    IF _runOneStep THEN
        _runOneStep := FALSE;
        RETURN;
    END_IF
END_IF

IF SUPER^.Step(765, TRUE, 'Step number 765') THEN
    SUPER^.StepCompleteWhen((_runOneStep OR _runAllSteps) AND _finishStep);

    IF _runOneStep THEN
        _runOneStep := FALSE;
        RETURN;
    END_IF
END_IF

IF SUPER^.Step(766, TRUE, 'Step number 766') THEN
    SUPER^.StepCompleteWhen((_runOneStep OR _runAllSteps) AND _finishStep);

    IF _runOneStep THEN
        _runOneStep := FALSE;
        RETURN;
    END_IF
END_IF

IF SUPER^.Step(767, TRUE, 'Step number 767') THEN
    SUPER^.StepCompleteWhen((_runOneStep OR _runAllSteps) AND _finishStep);

    IF _runOneStep THEN
        _runOneStep := FALSE;
        RETURN;
    END_IF
END_IF

IF SUPER^.Step(768, TRUE, 'Step number 768') THEN
    SUPER^.StepCompleteWhen((_runOneStep OR _runAllSteps) AND _finishStep);

    IF _runOneStep THEN
        _runOneStep := FALSE;
        RETURN;
    END_IF
END_IF

IF SUPER^.Step(769, TRUE, 'Step number 769') THEN
    SUPER^.StepCompleteWhen((_runOneStep OR _runAllSteps) AND _finishStep);

    IF _runOneStep THEN
        _runOneStep := FALSE;
        RETURN;
    END_IF
END_IF

IF SUPER^.Step(770, TRUE, 'Step number 770') THEN
    SUPER^.StepCompleteWhen((_runOneStep OR _runAllSteps) AND _finishStep);

    IF _runOneStep THEN
        _runOneStep := FALSE;
        RETURN;
    END_IF
END_IF

IF SUPER^.Step(771, TRUE, 'Step number 771') THEN
    SUPER^.StepCompleteWhen((_runOneStep OR _runAllSteps) AND _finishStep);

    IF _runOneStep THEN
        _runOneStep := FALSE;
        RETURN;
    END_IF
END_IF

IF SUPER^.Step(772, TRUE, 'Step number 772') THEN
    SUPER^.StepCompleteWhen((_runOneStep OR _runAllSteps) AND _finishStep);

    IF _runOneStep THEN
        _runOneStep := FALSE;
        RETURN;
    END_IF
END_IF

IF SUPER^.Step(773, TRUE, 'Step number 773') THEN
    SUPER^.StepCompleteWhen((_runOneStep OR _runAllSteps) AND _finishStep);

    IF _runOneStep THEN
        _runOneStep := FALSE;
        RETURN;
    END_IF
END_IF

IF SUPER^.Step(774, TRUE, 'Step number 774') THEN
    SUPER^.StepCompleteWhen((_runOneStep OR _runAllSteps) AND _finishStep);

    IF _runOneStep THEN
        _runOneStep := FALSE;
        RETURN;
    END_IF
END_IF

IF SUPER^.Step(775, TRUE, 'Step number 775') THEN
    SUPER^.StepCompleteWhen((_runOneStep OR _runAllSteps) AND _finishStep);

    IF _runOneStep THEN
        _runOneStep := FALSE;
        RETURN;
    END_IF
END_IF

IF SUPER^.Step(776, TRUE, 'Step number 776') THEN
    SUPER^.StepCompleteWhen((_runOneStep OR _runAllSteps) AND _finishStep);

    IF _runOneStep THEN
        _runOneStep := FALSE;
        RETURN;
    END_IF
END_IF

IF SUPER^.Step(777, TRUE, 'Step number 777') THEN
    SUPER^.StepCompleteWhen((_runOneStep OR _runAllSteps) AND _finishStep);

    IF _runOneStep THEN
        _runOneStep := FALSE;
        RETURN;
    END_IF
END_IF

IF SUPER^.Step(778, TRUE, 'Step number 778') THEN
    SUPER^.StepCompleteWhen((_runOneStep OR _runAllSteps) AND _finishStep);

    IF _runOneStep THEN
        _runOneStep := FALSE;
        RETURN;
    END_IF
END_IF

IF SUPER^.Step(779, TRUE, 'Step number 779') THEN
    SUPER^.StepCompleteWhen((_runOneStep OR _runAllSteps) AND _finishStep);

    IF _runOneStep THEN
        _runOneStep := FALSE;
        RETURN;
    END_IF
END_IF

IF SUPER^.Step(780, TRUE, 'Step number 780') THEN
    SUPER^.StepCompleteWhen((_runOneStep OR _runAllSteps) AND _finishStep);

    IF _runOneStep THEN
        _runOneStep := FALSE;
        RETURN;
    END_IF
END_IF

IF SUPER^.Step(781, TRUE, 'Step number 781') THEN
    SUPER^.StepCompleteWhen((_runOneStep OR _runAllSteps) AND _finishStep);

    IF _runOneStep THEN
        _runOneStep := FALSE;
        RETURN;
    END_IF
END_IF

IF SUPER^.Step(782, TRUE, 'Step number 782') THEN
    SUPER^.StepCompleteWhen((_runOneStep OR _runAllSteps) AND _finishStep);

    IF _runOneStep THEN
        _runOneStep := FALSE;
        RETURN;
    END_IF
END_IF

IF SUPER^.Step(783, TRUE, 'Step number 783') THEN
    SUPER^.StepCompleteWhen((_runOneStep OR _runAllSteps) AND _finishStep);

    IF _runOneStep THEN
        _runOneStep := FALSE;
        RETURN;
    END_IF
END_IF

IF SUPER^.Step(784, TRUE, 'Step number 784') THEN
    SUPER^.StepCompleteWhen((_runOneStep OR _runAllSteps) AND _finishStep);

    IF _runOneStep THEN
        _runOneStep := FALSE;
        RETURN;
    END_IF
END_IF

IF SUPER^.Step(785, TRUE, 'Step number 785') THEN
    SUPER^.StepCompleteWhen((_runOneStep OR _runAllSteps) AND _finishStep);

    IF _runOneStep THEN
        _runOneStep := FALSE;
        RETURN;
    END_IF
END_IF

IF SUPER^.Step(786, TRUE, 'Step number 786') THEN
    SUPER^.StepCompleteWhen((_runOneStep OR _runAllSteps) AND _finishStep);

    IF _runOneStep THEN
        _runOneStep := FALSE;
        RETURN;
    END_IF
END_IF

IF SUPER^.Step(787, TRUE, 'Step number 787') THEN
    SUPER^.StepCompleteWhen((_runOneStep OR _runAllSteps) AND _finishStep);

    IF _runOneStep THEN
        _runOneStep := FALSE;
        RETURN;
    END_IF
END_IF

IF SUPER^.Step(788, TRUE, 'Step number 788') THEN
    SUPER^.StepCompleteWhen((_runOneStep OR _runAllSteps) AND _finishStep);

    IF _runOneStep THEN
        _runOneStep := FALSE;
        RETURN;
    END_IF
END_IF

IF SUPER^.Step(789, TRUE, 'Step number 789') THEN
    SUPER^.StepCompleteWhen((_runOneStep OR _runAllSteps) AND _finishStep);

    IF _runOneStep THEN
        _runOneStep := FALSE;
        RETURN;
    END_IF
END_IF

IF SUPER^.Step(790, TRUE, 'Step number 790') THEN
    SUPER^.StepCompleteWhen((_runOneStep OR _runAllSteps) AND _finishStep);

    IF _runOneStep THEN
        _runOneStep := FALSE;
        RETURN;
    END_IF
END_IF

IF SUPER^.Step(791, TRUE, 'Step number 791') THEN
    SUPER^.StepCompleteWhen((_runOneStep OR _runAllSteps) AND _finishStep);

    IF _runOneStep THEN
        _runOneStep := FALSE;
        RETURN;
    END_IF
END_IF

IF SUPER^.Step(792, TRUE, 'Step number 792') THEN
    SUPER^.StepCompleteWhen((_runOneStep OR _runAllSteps) AND _finishStep);

    IF _runOneStep THEN
        _runOneStep := FALSE;
        RETURN;
    END_IF
END_IF

IF SUPER^.Step(793, TRUE, 'Step number 793') THEN
    SUPER^.StepCompleteWhen((_runOneStep OR _runAllSteps) AND _finishStep);

    IF _runOneStep THEN
        _runOneStep := FALSE;
        RETURN;
    END_IF
END_IF

IF SUPER^.Step(794, TRUE, 'Step number 794') THEN
    SUPER^.StepCompleteWhen((_runOneStep OR _runAllSteps) AND _finishStep);

    IF _runOneStep THEN
        _runOneStep := FALSE;
        RETURN;
    END_IF
END_IF

IF SUPER^.Step(795, TRUE, 'Step number 795') THEN
    SUPER^.StepCompleteWhen((_runOneStep OR _runAllSteps) AND _finishStep);

    IF _runOneStep THEN
        _runOneStep := FALSE;
        RETURN;
    END_IF
END_IF

IF SUPER^.Step(796, TRUE, 'Step number 796') THEN
    SUPER^.StepCompleteWhen((_runOneStep OR _runAllSteps) AND _finishStep);

    IF _runOneStep THEN
        _runOneStep := FALSE;
        RETURN;
    END_IF
END_IF

IF SUPER^.Step(797, TRUE, 'Step number 797') THEN
    SUPER^.StepCompleteWhen((_runOneStep OR _runAllSteps) AND _finishStep);

    IF _runOneStep THEN
        _runOneStep := FALSE;
        RETURN;
    END_IF
END_IF

IF SUPER^.Step(798, TRUE, 'Step number 798') THEN
    SUPER^.StepCompleteWhen((_runOneStep OR _runAllSteps) AND _finishStep);

    IF _runOneStep THEN
        _runOneStep := FALSE;
        RETURN;
    END_IF
END_IF

IF SUPER^.Step(799, TRUE, 'Step number 799') THEN
    SUPER^.StepCompleteWhen((_runOneStep OR _runAllSteps) AND _finishStep);

    IF _runOneStep THEN
        _runOneStep := FALSE;
        RETURN;
    END_IF
END_IF

IF SUPER^.Step(800, TRUE, 'Step number 800') THEN
    SUPER^.StepCompleteWhen((_runOneStep OR _runAllSteps) AND _finishStep);

    IF _runOneStep THEN
        _runOneStep := FALSE;
        RETURN;
    END_IF
END_IF

IF SUPER^.Step(801, TRUE, 'Step number 801') THEN
    SUPER^.StepCompleteWhen((_runOneStep OR _runAllSteps) AND _finishStep);

    IF _runOneStep THEN
        _runOneStep := FALSE;
        RETURN;
    END_IF
END_IF

IF SUPER^.Step(802, TRUE, 'Step number 802') THEN
    SUPER^.StepCompleteWhen((_runOneStep OR _runAllSteps) AND _finishStep);

    IF _runOneStep THEN
        _runOneStep := FALSE;
        RETURN;
    END_IF
END_IF

IF SUPER^.Step(803, TRUE, 'Step number 803') THEN
    SUPER^.StepCompleteWhen((_runOneStep OR _runAllSteps) AND _finishStep);

    IF _runOneStep THEN
        _runOneStep := FALSE;
        RETURN;
    END_IF
END_IF

IF SUPER^.Step(804, TRUE, 'Step number 804') THEN
    SUPER^.StepCompleteWhen((_runOneStep OR _runAllSteps) AND _finishStep);

    IF _runOneStep THEN
        _runOneStep := FALSE;
        RETURN;
    END_IF
END_IF

IF SUPER^.Step(805, TRUE, 'Step number 805') THEN
    SUPER^.StepCompleteWhen((_runOneStep OR _runAllSteps) AND _finishStep);

    IF _runOneStep THEN
        _runOneStep := FALSE;
        RETURN;
    END_IF
END_IF

IF SUPER^.Step(806, TRUE, 'Step number 806') THEN
    SUPER^.StepCompleteWhen((_runOneStep OR _runAllSteps) AND _finishStep);

    IF _runOneStep THEN
        _runOneStep := FALSE;
        RETURN;
    END_IF
END_IF

IF SUPER^.Step(807, TRUE, 'Step number 807') THEN
    SUPER^.StepCompleteWhen((_runOneStep OR _runAllSteps) AND _finishStep);

    IF _runOneStep THEN
        _runOneStep := FALSE;
        RETURN;
    END_IF
END_IF

IF SUPER^.Step(808, TRUE, 'Step number 808') THEN
    SUPER^.StepCompleteWhen((_runOneStep OR _runAllSteps) AND _finishStep);

    IF _runOneStep THEN
        _runOneStep := FALSE;
        RETURN;
    END_IF
END_IF

IF SUPER^.Step(809, TRUE, 'Step number 809') THEN
    SUPER^.StepCompleteWhen((_runOneStep OR _runAllSteps) AND _finishStep);

    IF _runOneStep THEN
        _runOneStep := FALSE;
        RETURN;
    END_IF
END_IF

IF SUPER^.Step(810, TRUE, 'Step number 810') THEN
    SUPER^.StepCompleteWhen((_runOneStep OR _runAllSteps) AND _finishStep);

    IF _runOneStep THEN
        _runOneStep := FALSE;
        RETURN;
    END_IF
END_IF

IF SUPER^.Step(811, TRUE, 'Step number 811') THEN
    SUPER^.StepCompleteWhen((_runOneStep OR _runAllSteps) AND _finishStep);

    IF _runOneStep THEN
        _runOneStep := FALSE;
        RETURN;
    END_IF
END_IF

IF SUPER^.Step(812, TRUE, 'Step number 812') THEN
    SUPER^.StepCompleteWhen((_runOneStep OR _runAllSteps) AND _finishStep);

    IF _runOneStep THEN
        _runOneStep := FALSE;
        RETURN;
    END_IF
END_IF

IF SUPER^.Step(813, TRUE, 'Step number 813') THEN
    SUPER^.StepCompleteWhen((_runOneStep OR _runAllSteps) AND _finishStep);

    IF _runOneStep THEN
        _runOneStep := FALSE;
        RETURN;
    END_IF
END_IF

IF SUPER^.Step(814, TRUE, 'Step number 814') THEN
    SUPER^.StepCompleteWhen((_runOneStep OR _runAllSteps) AND _finishStep);

    IF _runOneStep THEN
        _runOneStep := FALSE;
        RETURN;
    END_IF
END_IF

IF SUPER^.Step(815, TRUE, 'Step number 815') THEN
    SUPER^.StepCompleteWhen((_runOneStep OR _runAllSteps) AND _finishStep);

    IF _runOneStep THEN
        _runOneStep := FALSE;
        RETURN;
    END_IF
END_IF

IF SUPER^.Step(816, TRUE, 'Step number 816') THEN
    SUPER^.StepCompleteWhen((_runOneStep OR _runAllSteps) AND _finishStep);

    IF _runOneStep THEN
        _runOneStep := FALSE;
        RETURN;
    END_IF
END_IF

IF SUPER^.Step(817, TRUE, 'Step number 817') THEN
    SUPER^.StepCompleteWhen((_runOneStep OR _runAllSteps) AND _finishStep);

    IF _runOneStep THEN
        _runOneStep := FALSE;
        RETURN;
    END_IF
END_IF

IF SUPER^.Step(818, TRUE, 'Step number 818') THEN
    SUPER^.StepCompleteWhen((_runOneStep OR _runAllSteps) AND _finishStep);

    IF _runOneStep THEN
        _runOneStep := FALSE;
        RETURN;
    END_IF
END_IF

IF SUPER^.Step(819, TRUE, 'Step number 819') THEN
    SUPER^.StepCompleteWhen((_runOneStep OR _runAllSteps) AND _finishStep);

    IF _runOneStep THEN
        _runOneStep := FALSE;
        RETURN;
    END_IF
END_IF

IF SUPER^.Step(820, TRUE, 'Step number 820') THEN
    SUPER^.StepCompleteWhen((_runOneStep OR _runAllSteps) AND _finishStep);

    IF _runOneStep THEN
        _runOneStep := FALSE;
        RETURN;
    END_IF
END_IF

IF SUPER^.Step(821, TRUE, 'Step number 821') THEN
    SUPER^.StepCompleteWhen((_runOneStep OR _runAllSteps) AND _finishStep);

    IF _runOneStep THEN
        _runOneStep := FALSE;
        RETURN;
    END_IF
END_IF

IF SUPER^.Step(822, TRUE, 'Step number 822') THEN
    SUPER^.StepCompleteWhen((_runOneStep OR _runAllSteps) AND _finishStep);

    IF _runOneStep THEN
        _runOneStep := FALSE;
        RETURN;
    END_IF
END_IF

IF SUPER^.Step(823, TRUE, 'Step number 823') THEN
    SUPER^.StepCompleteWhen((_runOneStep OR _runAllSteps) AND _finishStep);

    IF _runOneStep THEN
        _runOneStep := FALSE;
        RETURN;
    END_IF
END_IF

IF SUPER^.Step(824, TRUE, 'Step number 824') THEN
    SUPER^.StepCompleteWhen((_runOneStep OR _runAllSteps) AND _finishStep);

    IF _runOneStep THEN
        _runOneStep := FALSE;
        RETURN;
    END_IF
END_IF

IF SUPER^.Step(825, TRUE, 'Step number 825') THEN
    SUPER^.StepCompleteWhen((_runOneStep OR _runAllSteps) AND _finishStep);

    IF _runOneStep THEN
        _runOneStep := FALSE;
        RETURN;
    END_IF
END_IF

IF SUPER^.Step(826, TRUE, 'Step number 826') THEN
    SUPER^.StepCompleteWhen((_runOneStep OR _runAllSteps) AND _finishStep);

    IF _runOneStep THEN
        _runOneStep := FALSE;
        RETURN;
    END_IF
END_IF

IF SUPER^.Step(827, TRUE, 'Step number 827') THEN
    SUPER^.StepCompleteWhen((_runOneStep OR _runAllSteps) AND _finishStep);

    IF _runOneStep THEN
        _runOneStep := FALSE;
        RETURN;
    END_IF
END_IF

IF SUPER^.Step(828, TRUE, 'Step number 828') THEN
    SUPER^.StepCompleteWhen((_runOneStep OR _runAllSteps) AND _finishStep);

    IF _runOneStep THEN
        _runOneStep := FALSE;
        RETURN;
    END_IF
END_IF

IF SUPER^.Step(829, TRUE, 'Step number 829') THEN
    SUPER^.StepCompleteWhen((_runOneStep OR _runAllSteps) AND _finishStep);

    IF _runOneStep THEN
        _runOneStep := FALSE;
        RETURN;
    END_IF
END_IF

IF SUPER^.Step(830, TRUE, 'Step number 830') THEN
    SUPER^.StepCompleteWhen((_runOneStep OR _runAllSteps) AND _finishStep);

    IF _runOneStep THEN
        _runOneStep := FALSE;
        RETURN;
    END_IF
END_IF

IF SUPER^.Step(831, TRUE, 'Step number 831') THEN
    SUPER^.StepCompleteWhen((_runOneStep OR _runAllSteps) AND _finishStep);

    IF _runOneStep THEN
        _runOneStep := FALSE;
        RETURN;
    END_IF
END_IF

IF SUPER^.Step(832, TRUE, 'Step number 832') THEN
    SUPER^.StepCompleteWhen((_runOneStep OR _runAllSteps) AND _finishStep);

    IF _runOneStep THEN
        _runOneStep := FALSE;
        RETURN;
    END_IF
END_IF

IF SUPER^.Step(833, TRUE, 'Step number 833') THEN
    SUPER^.StepCompleteWhen((_runOneStep OR _runAllSteps) AND _finishStep);

    IF _runOneStep THEN
        _runOneStep := FALSE;
        RETURN;
    END_IF
END_IF

IF SUPER^.Step(834, TRUE, 'Step number 834') THEN
    SUPER^.StepCompleteWhen((_runOneStep OR _runAllSteps) AND _finishStep);

    IF _runOneStep THEN
        _runOneStep := FALSE;
        RETURN;
    END_IF
END_IF

IF SUPER^.Step(835, TRUE, 'Step number 835') THEN
    SUPER^.StepCompleteWhen((_runOneStep OR _runAllSteps) AND _finishStep);

    IF _runOneStep THEN
        _runOneStep := FALSE;
        RETURN;
    END_IF
END_IF

IF SUPER^.Step(836, TRUE, 'Step number 836') THEN
    SUPER^.StepCompleteWhen((_runOneStep OR _runAllSteps) AND _finishStep);

    IF _runOneStep THEN
        _runOneStep := FALSE;
        RETURN;
    END_IF
END_IF

IF SUPER^.Step(837, TRUE, 'Step number 837') THEN
    SUPER^.StepCompleteWhen((_runOneStep OR _runAllSteps) AND _finishStep);

    IF _runOneStep THEN
        _runOneStep := FALSE;
        RETURN;
    END_IF
END_IF

IF SUPER^.Step(838, TRUE, 'Step number 838') THEN
    SUPER^.StepCompleteWhen((_runOneStep OR _runAllSteps) AND _finishStep);

    IF _runOneStep THEN
        _runOneStep := FALSE;
        RETURN;
    END_IF
END_IF

IF SUPER^.Step(839, TRUE, 'Step number 839') THEN
    SUPER^.StepCompleteWhen((_runOneStep OR _runAllSteps) AND _finishStep);

    IF _runOneStep THEN
        _runOneStep := FALSE;
        RETURN;
    END_IF
END_IF

IF SUPER^.Step(840, TRUE, 'Step number 840') THEN
    SUPER^.StepCompleteWhen((_runOneStep OR _runAllSteps) AND _finishStep);

    IF _runOneStep THEN
        _runOneStep := FALSE;
        RETURN;
    END_IF
END_IF

IF SUPER^.Step(841, TRUE, 'Step number 841') THEN
    SUPER^.StepCompleteWhen((_runOneStep OR _runAllSteps) AND _finishStep);

    IF _runOneStep THEN
        _runOneStep := FALSE;
        RETURN;
    END_IF
END_IF

IF SUPER^.Step(842, TRUE, 'Step number 842') THEN
    SUPER^.StepCompleteWhen((_runOneStep OR _runAllSteps) AND _finishStep);

    IF _runOneStep THEN
        _runOneStep := FALSE;
        RETURN;
    END_IF
END_IF

IF SUPER^.Step(843, TRUE, 'Step number 843') THEN
    SUPER^.StepCompleteWhen((_runOneStep OR _runAllSteps) AND _finishStep);

    IF _runOneStep THEN
        _runOneStep := FALSE;
        RETURN;
    END_IF
END_IF

IF SUPER^.Step(844, TRUE, 'Step number 844') THEN
    SUPER^.StepCompleteWhen((_runOneStep OR _runAllSteps) AND _finishStep);

    IF _runOneStep THEN
        _runOneStep := FALSE;
        RETURN;
    END_IF
END_IF

IF SUPER^.Step(845, TRUE, 'Step number 845') THEN
    SUPER^.StepCompleteWhen((_runOneStep OR _runAllSteps) AND _finishStep);

    IF _runOneStep THEN
        _runOneStep := FALSE;
        RETURN;
    END_IF
END_IF

IF SUPER^.Step(846, TRUE, 'Step number 846') THEN
    SUPER^.StepCompleteWhen((_runOneStep OR _runAllSteps) AND _finishStep);

    IF _runOneStep THEN
        _runOneStep := FALSE;
        RETURN;
    END_IF
END_IF

IF SUPER^.Step(847, TRUE, 'Step number 847') THEN
    SUPER^.StepCompleteWhen((_runOneStep OR _runAllSteps) AND _finishStep);

    IF _runOneStep THEN
        _runOneStep := FALSE;
        RETURN;
    END_IF
END_IF

IF SUPER^.Step(848, TRUE, 'Step number 848') THEN
    SUPER^.StepCompleteWhen((_runOneStep OR _runAllSteps) AND _finishStep);

    IF _runOneStep THEN
        _runOneStep := FALSE;
        RETURN;
    END_IF
END_IF

IF SUPER^.Step(849, TRUE, 'Step number 849') THEN
    SUPER^.StepCompleteWhen((_runOneStep OR _runAllSteps) AND _finishStep);

    IF _runOneStep THEN
        _runOneStep := FALSE;
        RETURN;
    END_IF
END_IF

IF SUPER^.Step(850, TRUE, 'Step number 850') THEN
    SUPER^.StepCompleteWhen((_runOneStep OR _runAllSteps) AND _finishStep);

    IF _runOneStep THEN
        _runOneStep := FALSE;
        RETURN;
    END_IF
END_IF

IF SUPER^.Step(851, TRUE, 'Step number 851') THEN
    SUPER^.StepCompleteWhen((_runOneStep OR _runAllSteps) AND _finishStep);

    IF _runOneStep THEN
        _runOneStep := FALSE;
        RETURN;
    END_IF
END_IF

IF SUPER^.Step(852, TRUE, 'Step number 852') THEN
    SUPER^.StepCompleteWhen((_runOneStep OR _runAllSteps) AND _finishStep);

    IF _runOneStep THEN
        _runOneStep := FALSE;
        RETURN;
    END_IF
END_IF

IF SUPER^.Step(853, TRUE, 'Step number 853') THEN
    SUPER^.StepCompleteWhen((_runOneStep OR _runAllSteps) AND _finishStep);

    IF _runOneStep THEN
        _runOneStep := FALSE;
        RETURN;
    END_IF
END_IF

IF SUPER^.Step(854, TRUE, 'Step number 854') THEN
    SUPER^.StepCompleteWhen((_runOneStep OR _runAllSteps) AND _finishStep);

    IF _runOneStep THEN
        _runOneStep := FALSE;
        RETURN;
    END_IF
END_IF

IF SUPER^.Step(855, TRUE, 'Step number 855') THEN
    SUPER^.StepCompleteWhen((_runOneStep OR _runAllSteps) AND _finishStep);

    IF _runOneStep THEN
        _runOneStep := FALSE;
        RETURN;
    END_IF
END_IF

IF SUPER^.Step(856, TRUE, 'Step number 856') THEN
    SUPER^.StepCompleteWhen((_runOneStep OR _runAllSteps) AND _finishStep);

    IF _runOneStep THEN
        _runOneStep := FALSE;
        RETURN;
    END_IF
END_IF

IF SUPER^.Step(857, TRUE, 'Step number 857') THEN
    SUPER^.StepCompleteWhen((_runOneStep OR _runAllSteps) AND _finishStep);

    IF _runOneStep THEN
        _runOneStep := FALSE;
        RETURN;
    END_IF
END_IF

IF SUPER^.Step(858, TRUE, 'Step number 858') THEN
    SUPER^.StepCompleteWhen((_runOneStep OR _runAllSteps) AND _finishStep);

    IF _runOneStep THEN
        _runOneStep := FALSE;
        RETURN;
    END_IF
END_IF

IF SUPER^.Step(859, TRUE, 'Step number 859') THEN
    SUPER^.StepCompleteWhen((_runOneStep OR _runAllSteps) AND _finishStep);

    IF _runOneStep THEN
        _runOneStep := FALSE;
        RETURN;
    END_IF
END_IF

IF SUPER^.Step(860, TRUE, 'Step number 860') THEN
    SUPER^.StepCompleteWhen((_runOneStep OR _runAllSteps) AND _finishStep);

    IF _runOneStep THEN
        _runOneStep := FALSE;
        RETURN;
    END_IF
END_IF

IF SUPER^.Step(861, TRUE, 'Step number 861') THEN
    SUPER^.StepCompleteWhen((_runOneStep OR _runAllSteps) AND _finishStep);

    IF _runOneStep THEN
        _runOneStep := FALSE;
        RETURN;
    END_IF
END_IF

IF SUPER^.Step(862, TRUE, 'Step number 862') THEN
    SUPER^.StepCompleteWhen((_runOneStep OR _runAllSteps) AND _finishStep);

    IF _runOneStep THEN
        _runOneStep := FALSE;
        RETURN;
    END_IF
END_IF

IF SUPER^.Step(863, TRUE, 'Step number 863') THEN
    SUPER^.StepCompleteWhen((_runOneStep OR _runAllSteps) AND _finishStep);

    IF _runOneStep THEN
        _runOneStep := FALSE;
        RETURN;
    END_IF
END_IF

IF SUPER^.Step(864, TRUE, 'Step number 864') THEN
    SUPER^.StepCompleteWhen((_runOneStep OR _runAllSteps) AND _finishStep);

    IF _runOneStep THEN
        _runOneStep := FALSE;
        RETURN;
    END_IF
END_IF

IF SUPER^.Step(865, TRUE, 'Step number 865') THEN
    SUPER^.StepCompleteWhen((_runOneStep OR _runAllSteps) AND _finishStep);

    IF _runOneStep THEN
        _runOneStep := FALSE;
        RETURN;
    END_IF
END_IF

IF SUPER^.Step(866, TRUE, 'Step number 866') THEN
    SUPER^.StepCompleteWhen((_runOneStep OR _runAllSteps) AND _finishStep);

    IF _runOneStep THEN
        _runOneStep := FALSE;
        RETURN;
    END_IF
END_IF

IF SUPER^.Step(867, TRUE, 'Step number 867') THEN
    SUPER^.StepCompleteWhen((_runOneStep OR _runAllSteps) AND _finishStep);

    IF _runOneStep THEN
        _runOneStep := FALSE;
        RETURN;
    END_IF
END_IF

IF SUPER^.Step(868, TRUE, 'Step number 868') THEN
    SUPER^.StepCompleteWhen((_runOneStep OR _runAllSteps) AND _finishStep);

    IF _runOneStep THEN
        _runOneStep := FALSE;
        RETURN;
    END_IF
END_IF

IF SUPER^.Step(869, TRUE, 'Step number 869') THEN
    SUPER^.StepCompleteWhen((_runOneStep OR _runAllSteps) AND _finishStep);

    IF _runOneStep THEN
        _runOneStep := FALSE;
        RETURN;
    END_IF
END_IF

IF SUPER^.Step(870, TRUE, 'Step number 870') THEN
    SUPER^.StepCompleteWhen((_runOneStep OR _runAllSteps) AND _finishStep);

    IF _runOneStep THEN
        _runOneStep := FALSE;
        RETURN;
    END_IF
END_IF

IF SUPER^.Step(871, TRUE, 'Step number 871') THEN
    SUPER^.StepCompleteWhen((_runOneStep OR _runAllSteps) AND _finishStep);

    IF _runOneStep THEN
        _runOneStep := FALSE;
        RETURN;
    END_IF
END_IF

IF SUPER^.Step(872, TRUE, 'Step number 872') THEN
    SUPER^.StepCompleteWhen((_runOneStep OR _runAllSteps) AND _finishStep);

    IF _runOneStep THEN
        _runOneStep := FALSE;
        RETURN;
    END_IF
END_IF

IF SUPER^.Step(873, TRUE, 'Step number 873') THEN
    SUPER^.StepCompleteWhen((_runOneStep OR _runAllSteps) AND _finishStep);

    IF _runOneStep THEN
        _runOneStep := FALSE;
        RETURN;
    END_IF
END_IF

IF SUPER^.Step(874, TRUE, 'Step number 874') THEN
    SUPER^.StepCompleteWhen((_runOneStep OR _runAllSteps) AND _finishStep);

    IF _runOneStep THEN
        _runOneStep := FALSE;
        RETURN;
    END_IF
END_IF

IF SUPER^.Step(875, TRUE, 'Step number 875') THEN
    SUPER^.StepCompleteWhen((_runOneStep OR _runAllSteps) AND _finishStep);

    IF _runOneStep THEN
        _runOneStep := FALSE;
        RETURN;
    END_IF
END_IF

IF SUPER^.Step(876, TRUE, 'Step number 876') THEN
    SUPER^.StepCompleteWhen((_runOneStep OR _runAllSteps) AND _finishStep);

    IF _runOneStep THEN
        _runOneStep := FALSE;
        RETURN;
    END_IF
END_IF

IF SUPER^.Step(877, TRUE, 'Step number 877') THEN
    SUPER^.StepCompleteWhen((_runOneStep OR _runAllSteps) AND _finishStep);

    IF _runOneStep THEN
        _runOneStep := FALSE;
        RETURN;
    END_IF
END_IF

IF SUPER^.Step(878, TRUE, 'Step number 878') THEN
    SUPER^.StepCompleteWhen((_runOneStep OR _runAllSteps) AND _finishStep);

    IF _runOneStep THEN
        _runOneStep := FALSE;
        RETURN;
    END_IF
END_IF

IF SUPER^.Step(879, TRUE, 'Step number 879') THEN
    SUPER^.StepCompleteWhen((_runOneStep OR _runAllSteps) AND _finishStep);

    IF _runOneStep THEN
        _runOneStep := FALSE;
        RETURN;
    END_IF
END_IF

IF SUPER^.Step(880, TRUE, 'Step number 880') THEN
    SUPER^.StepCompleteWhen((_runOneStep OR _runAllSteps) AND _finishStep);

    IF _runOneStep THEN
        _runOneStep := FALSE;
        RETURN;
    END_IF
END_IF

IF SUPER^.Step(881, TRUE, 'Step number 881') THEN
    SUPER^.StepCompleteWhen((_runOneStep OR _runAllSteps) AND _finishStep);

    IF _runOneStep THEN
        _runOneStep := FALSE;
        RETURN;
    END_IF
END_IF

IF SUPER^.Step(882, TRUE, 'Step number 882') THEN
    SUPER^.StepCompleteWhen((_runOneStep OR _runAllSteps) AND _finishStep);

    IF _runOneStep THEN
        _runOneStep := FALSE;
        RETURN;
    END_IF
END_IF

IF SUPER^.Step(883, TRUE, 'Step number 883') THEN
    SUPER^.StepCompleteWhen((_runOneStep OR _runAllSteps) AND _finishStep);

    IF _runOneStep THEN
        _runOneStep := FALSE;
        RETURN;
    END_IF
END_IF

IF SUPER^.Step(884, TRUE, 'Step number 884') THEN
    SUPER^.StepCompleteWhen((_runOneStep OR _runAllSteps) AND _finishStep);

    IF _runOneStep THEN
        _runOneStep := FALSE;
        RETURN;
    END_IF
END_IF

IF SUPER^.Step(885, TRUE, 'Step number 885') THEN
    SUPER^.StepCompleteWhen((_runOneStep OR _runAllSteps) AND _finishStep);

    IF _runOneStep THEN
        _runOneStep := FALSE;
        RETURN;
    END_IF
END_IF

IF SUPER^.Step(886, TRUE, 'Step number 886') THEN
    SUPER^.StepCompleteWhen((_runOneStep OR _runAllSteps) AND _finishStep);

    IF _runOneStep THEN
        _runOneStep := FALSE;
        RETURN;
    END_IF
END_IF

IF SUPER^.Step(887, TRUE, 'Step number 887') THEN
    SUPER^.StepCompleteWhen((_runOneStep OR _runAllSteps) AND _finishStep);

    IF _runOneStep THEN
        _runOneStep := FALSE;
        RETURN;
    END_IF
END_IF

IF SUPER^.Step(888, TRUE, 'Step number 888') THEN
    SUPER^.StepCompleteWhen((_runOneStep OR _runAllSteps) AND _finishStep);

    IF _runOneStep THEN
        _runOneStep := FALSE;
        RETURN;
    END_IF
END_IF

IF SUPER^.Step(889, TRUE, 'Step number 889') THEN
    SUPER^.StepCompleteWhen((_runOneStep OR _runAllSteps) AND _finishStep);

    IF _runOneStep THEN
        _runOneStep := FALSE;
        RETURN;
    END_IF
END_IF

IF SUPER^.Step(890, TRUE, 'Step number 890') THEN
    SUPER^.StepCompleteWhen((_runOneStep OR _runAllSteps) AND _finishStep);

    IF _runOneStep THEN
        _runOneStep := FALSE;
        RETURN;
    END_IF
END_IF

IF SUPER^.Step(891, TRUE, 'Step number 891') THEN
    SUPER^.StepCompleteWhen((_runOneStep OR _runAllSteps) AND _finishStep);

    IF _runOneStep THEN
        _runOneStep := FALSE;
        RETURN;
    END_IF
END_IF

IF SUPER^.Step(892, TRUE, 'Step number 892') THEN
    SUPER^.StepCompleteWhen((_runOneStep OR _runAllSteps) AND _finishStep);

    IF _runOneStep THEN
        _runOneStep := FALSE;
        RETURN;
    END_IF
END_IF

IF SUPER^.Step(893, TRUE, 'Step number 893') THEN
    SUPER^.StepCompleteWhen((_runOneStep OR _runAllSteps) AND _finishStep);

    IF _runOneStep THEN
        _runOneStep := FALSE;
        RETURN;
    END_IF
END_IF

IF SUPER^.Step(894, TRUE, 'Step number 894') THEN
    SUPER^.StepCompleteWhen((_runOneStep OR _runAllSteps) AND _finishStep);

    IF _runOneStep THEN
        _runOneStep := FALSE;
        RETURN;
    END_IF
END_IF

IF SUPER^.Step(895, TRUE, 'Step number 895') THEN
    SUPER^.StepCompleteWhen((_runOneStep OR _runAllSteps) AND _finishStep);

    IF _runOneStep THEN
        _runOneStep := FALSE;
        RETURN;
    END_IF
END_IF

IF SUPER^.Step(896, TRUE, 'Step number 896') THEN
    SUPER^.StepCompleteWhen((_runOneStep OR _runAllSteps) AND _finishStep);

    IF _runOneStep THEN
        _runOneStep := FALSE;
        RETURN;
    END_IF
END_IF

IF SUPER^.Step(897, TRUE, 'Step number 897') THEN
    SUPER^.StepCompleteWhen((_runOneStep OR _runAllSteps) AND _finishStep);

    IF _runOneStep THEN
        _runOneStep := FALSE;
        RETURN;
    END_IF
END_IF

IF SUPER^.Step(898, TRUE, 'Step number 898') THEN
    SUPER^.StepCompleteWhen((_runOneStep OR _runAllSteps) AND _finishStep);

    IF _runOneStep THEN
        _runOneStep := FALSE;
        RETURN;
    END_IF
END_IF

IF SUPER^.Step(899, TRUE, 'Step number 899') THEN
    SUPER^.StepCompleteWhen((_runOneStep OR _runAllSteps) AND _finishStep);

    IF _runOneStep THEN
        _runOneStep := FALSE;
        RETURN;
    END_IF
END_IF

IF SUPER^.Step(900, TRUE, 'Step number 900') THEN
    SUPER^.StepCompleteWhen((_runOneStep OR _runAllSteps) AND _finishStep);

    IF _runOneStep THEN
        _runOneStep := FALSE;
        RETURN;
    END_IF
END_IF

IF SUPER^.Step(901, TRUE, 'Step number 901') THEN
    SUPER^.StepCompleteWhen((_runOneStep OR _runAllSteps) AND _finishStep);

    IF _runOneStep THEN
        _runOneStep := FALSE;
        RETURN;
    END_IF
END_IF

IF SUPER^.Step(902, TRUE, 'Step number 902') THEN
    SUPER^.StepCompleteWhen((_runOneStep OR _runAllSteps) AND _finishStep);

    IF _runOneStep THEN
        _runOneStep := FALSE;
        RETURN;
    END_IF
END_IF

IF SUPER^.Step(903, TRUE, 'Step number 903') THEN
    SUPER^.StepCompleteWhen((_runOneStep OR _runAllSteps) AND _finishStep);

    IF _runOneStep THEN
        _runOneStep := FALSE;
        RETURN;
    END_IF
END_IF

IF SUPER^.Step(904, TRUE, 'Step number 904') THEN
    SUPER^.StepCompleteWhen((_runOneStep OR _runAllSteps) AND _finishStep);

    IF _runOneStep THEN
        _runOneStep := FALSE;
        RETURN;
    END_IF
END_IF

IF SUPER^.Step(905, TRUE, 'Step number 905') THEN
    SUPER^.StepCompleteWhen((_runOneStep OR _runAllSteps) AND _finishStep);

    IF _runOneStep THEN
        _runOneStep := FALSE;
        RETURN;
    END_IF
END_IF

IF SUPER^.Step(906, TRUE, 'Step number 906') THEN
    SUPER^.StepCompleteWhen((_runOneStep OR _runAllSteps) AND _finishStep);

    IF _runOneStep THEN
        _runOneStep := FALSE;
        RETURN;
    END_IF
END_IF

IF SUPER^.Step(907, TRUE, 'Step number 907') THEN
    SUPER^.StepCompleteWhen((_runOneStep OR _runAllSteps) AND _finishStep);

    IF _runOneStep THEN
        _runOneStep := FALSE;
        RETURN;
    END_IF
END_IF

IF SUPER^.Step(908, TRUE, 'Step number 908') THEN
    SUPER^.StepCompleteWhen((_runOneStep OR _runAllSteps) AND _finishStep);

    IF _runOneStep THEN
        _runOneStep := FALSE;
        RETURN;
    END_IF
END_IF

IF SUPER^.Step(909, TRUE, 'Step number 909') THEN
    SUPER^.StepCompleteWhen((_runOneStep OR _runAllSteps) AND _finishStep);

    IF _runOneStep THEN
        _runOneStep := FALSE;
        RETURN;
    END_IF
END_IF

IF SUPER^.Step(910, TRUE, 'Step number 910') THEN
    SUPER^.StepCompleteWhen((_runOneStep OR _runAllSteps) AND _finishStep);

    IF _runOneStep THEN
        _runOneStep := FALSE;
        RETURN;
    END_IF
END_IF

IF SUPER^.Step(911, TRUE, 'Step number 911') THEN
    SUPER^.StepCompleteWhen((_runOneStep OR _runAllSteps) AND _finishStep);

    IF _runOneStep THEN
        _runOneStep := FALSE;
        RETURN;
    END_IF
END_IF

IF SUPER^.Step(912, TRUE, 'Step number 912') THEN
    SUPER^.StepCompleteWhen((_runOneStep OR _runAllSteps) AND _finishStep);

    IF _runOneStep THEN
        _runOneStep := FALSE;
        RETURN;
    END_IF
END_IF

IF SUPER^.Step(913, TRUE, 'Step number 913') THEN
    SUPER^.StepCompleteWhen((_runOneStep OR _runAllSteps) AND _finishStep);

    IF _runOneStep THEN
        _runOneStep := FALSE;
        RETURN;
    END_IF
END_IF

IF SUPER^.Step(914, TRUE, 'Step number 914') THEN
    SUPER^.StepCompleteWhen((_runOneStep OR _runAllSteps) AND _finishStep);

    IF _runOneStep THEN
        _runOneStep := FALSE;
        RETURN;
    END_IF
END_IF

IF SUPER^.Step(915, TRUE, 'Step number 915') THEN
    SUPER^.StepCompleteWhen((_runOneStep OR _runAllSteps) AND _finishStep);

    IF _runOneStep THEN
        _runOneStep := FALSE;
        RETURN;
    END_IF
END_IF

IF SUPER^.Step(916, TRUE, 'Step number 916') THEN
    SUPER^.StepCompleteWhen((_runOneStep OR _runAllSteps) AND _finishStep);

    IF _runOneStep THEN
        _runOneStep := FALSE;
        RETURN;
    END_IF
END_IF

IF SUPER^.Step(917, TRUE, 'Step number 917') THEN
    SUPER^.StepCompleteWhen((_runOneStep OR _runAllSteps) AND _finishStep);

    IF _runOneStep THEN
        _runOneStep := FALSE;
        RETURN;
    END_IF
END_IF

IF SUPER^.Step(918, TRUE, 'Step number 918') THEN
    SUPER^.StepCompleteWhen((_runOneStep OR _runAllSteps) AND _finishStep);

    IF _runOneStep THEN
        _runOneStep := FALSE;
        RETURN;
    END_IF
END_IF

IF SUPER^.Step(919, TRUE, 'Step number 919') THEN
    SUPER^.StepCompleteWhen((_runOneStep OR _runAllSteps) AND _finishStep);

    IF _runOneStep THEN
        _runOneStep := FALSE;
        RETURN;
    END_IF
END_IF

IF SUPER^.Step(920, TRUE, 'Step number 920') THEN
    SUPER^.StepCompleteWhen((_runOneStep OR _runAllSteps) AND _finishStep);

    IF _runOneStep THEN
        _runOneStep := FALSE;
        RETURN;
    END_IF
END_IF

IF SUPER^.Step(921, TRUE, 'Step number 921') THEN
    SUPER^.StepCompleteWhen((_runOneStep OR _runAllSteps) AND _finishStep);

    IF _runOneStep THEN
        _runOneStep := FALSE;
        RETURN;
    END_IF
END_IF

IF SUPER^.Step(922, TRUE, 'Step number 922') THEN
    SUPER^.StepCompleteWhen((_runOneStep OR _runAllSteps) AND _finishStep);

    IF _runOneStep THEN
        _runOneStep := FALSE;
        RETURN;
    END_IF
END_IF

IF SUPER^.Step(923, TRUE, 'Step number 923') THEN
    SUPER^.StepCompleteWhen((_runOneStep OR _runAllSteps) AND _finishStep);

    IF _runOneStep THEN
        _runOneStep := FALSE;
        RETURN;
    END_IF
END_IF

IF SUPER^.Step(924, TRUE, 'Step number 924') THEN
    SUPER^.StepCompleteWhen((_runOneStep OR _runAllSteps) AND _finishStep);

    IF _runOneStep THEN
        _runOneStep := FALSE;
        RETURN;
    END_IF
END_IF

IF SUPER^.Step(925, TRUE, 'Step number 925') THEN
    SUPER^.StepCompleteWhen((_runOneStep OR _runAllSteps) AND _finishStep);

    IF _runOneStep THEN
        _runOneStep := FALSE;
        RETURN;
    END_IF
END_IF

IF SUPER^.Step(926, TRUE, 'Step number 926') THEN
    SUPER^.StepCompleteWhen((_runOneStep OR _runAllSteps) AND _finishStep);

    IF _runOneStep THEN
        _runOneStep := FALSE;
        RETURN;
    END_IF
END_IF

IF SUPER^.Step(927, TRUE, 'Step number 927') THEN
    SUPER^.StepCompleteWhen((_runOneStep OR _runAllSteps) AND _finishStep);

    IF _runOneStep THEN
        _runOneStep := FALSE;
        RETURN;
    END_IF
END_IF

IF SUPER^.Step(928, TRUE, 'Step number 928') THEN
    SUPER^.StepCompleteWhen((_runOneStep OR _runAllSteps) AND _finishStep);

    IF _runOneStep THEN
        _runOneStep := FALSE;
        RETURN;
    END_IF
END_IF

IF SUPER^.Step(929, TRUE, 'Step number 929') THEN
    SUPER^.StepCompleteWhen((_runOneStep OR _runAllSteps) AND _finishStep);

    IF _runOneStep THEN
        _runOneStep := FALSE;
        RETURN;
    END_IF
END_IF

IF SUPER^.Step(930, TRUE, 'Step number 930') THEN
    SUPER^.StepCompleteWhen((_runOneStep OR _runAllSteps) AND _finishStep);

    IF _runOneStep THEN
        _runOneStep := FALSE;
        RETURN;
    END_IF
END_IF

IF SUPER^.Step(931, TRUE, 'Step number 931') THEN
    SUPER^.StepCompleteWhen((_runOneStep OR _runAllSteps) AND _finishStep);

    IF _runOneStep THEN
        _runOneStep := FALSE;
        RETURN;
    END_IF
END_IF

IF SUPER^.Step(932, TRUE, 'Step number 932') THEN
    SUPER^.StepCompleteWhen((_runOneStep OR _runAllSteps) AND _finishStep);

    IF _runOneStep THEN
        _runOneStep := FALSE;
        RETURN;
    END_IF
END_IF

IF SUPER^.Step(933, TRUE, 'Step number 933') THEN
    SUPER^.StepCompleteWhen((_runOneStep OR _runAllSteps) AND _finishStep);

    IF _runOneStep THEN
        _runOneStep := FALSE;
        RETURN;
    END_IF
END_IF

IF SUPER^.Step(934, TRUE, 'Step number 934') THEN
    SUPER^.StepCompleteWhen((_runOneStep OR _runAllSteps) AND _finishStep);

    IF _runOneStep THEN
        _runOneStep := FALSE;
        RETURN;
    END_IF
END_IF

IF SUPER^.Step(935, TRUE, 'Step number 935') THEN
    SUPER^.StepCompleteWhen((_runOneStep OR _runAllSteps) AND _finishStep);

    IF _runOneStep THEN
        _runOneStep := FALSE;
        RETURN;
    END_IF
END_IF

IF SUPER^.Step(936, TRUE, 'Step number 936') THEN
    SUPER^.StepCompleteWhen((_runOneStep OR _runAllSteps) AND _finishStep);

    IF _runOneStep THEN
        _runOneStep := FALSE;
        RETURN;
    END_IF
END_IF

IF SUPER^.Step(937, TRUE, 'Step number 937') THEN
    SUPER^.StepCompleteWhen((_runOneStep OR _runAllSteps) AND _finishStep);

    IF _runOneStep THEN
        _runOneStep := FALSE;
        RETURN;
    END_IF
END_IF

IF SUPER^.Step(938, TRUE, 'Step number 938') THEN
    SUPER^.StepCompleteWhen((_runOneStep OR _runAllSteps) AND _finishStep);

    IF _runOneStep THEN
        _runOneStep := FALSE;
        RETURN;
    END_IF
END_IF

IF SUPER^.Step(939, TRUE, 'Step number 939') THEN
    SUPER^.StepCompleteWhen((_runOneStep OR _runAllSteps) AND _finishStep);

    IF _runOneStep THEN
        _runOneStep := FALSE;
        RETURN;
    END_IF
END_IF

IF SUPER^.Step(940, TRUE, 'Step number 940') THEN
    SUPER^.StepCompleteWhen((_runOneStep OR _runAllSteps) AND _finishStep);

    IF _runOneStep THEN
        _runOneStep := FALSE;
        RETURN;
    END_IF
END_IF

IF SUPER^.Step(941, TRUE, 'Step number 941') THEN
    SUPER^.StepCompleteWhen((_runOneStep OR _runAllSteps) AND _finishStep);

    IF _runOneStep THEN
        _runOneStep := FALSE;
        RETURN;
    END_IF
END_IF

IF SUPER^.Step(942, TRUE, 'Step number 942') THEN
    SUPER^.StepCompleteWhen((_runOneStep OR _runAllSteps) AND _finishStep);

    IF _runOneStep THEN
        _runOneStep := FALSE;
        RETURN;
    END_IF
END_IF

IF SUPER^.Step(943, TRUE, 'Step number 943') THEN
    SUPER^.StepCompleteWhen((_runOneStep OR _runAllSteps) AND _finishStep);

    IF _runOneStep THEN
        _runOneStep := FALSE;
        RETURN;
    END_IF
END_IF

IF SUPER^.Step(944, TRUE, 'Step number 944') THEN
    SUPER^.StepCompleteWhen((_runOneStep OR _runAllSteps) AND _finishStep);

    IF _runOneStep THEN
        _runOneStep := FALSE;
        RETURN;
    END_IF
END_IF

IF SUPER^.Step(945, TRUE, 'Step number 945') THEN
    SUPER^.StepCompleteWhen((_runOneStep OR _runAllSteps) AND _finishStep);

    IF _runOneStep THEN
        _runOneStep := FALSE;
        RETURN;
    END_IF
END_IF

IF SUPER^.Step(946, TRUE, 'Step number 946') THEN
    SUPER^.StepCompleteWhen((_runOneStep OR _runAllSteps) AND _finishStep);

    IF _runOneStep THEN
        _runOneStep := FALSE;
        RETURN;
    END_IF
END_IF

IF SUPER^.Step(947, TRUE, 'Step number 947') THEN
    SUPER^.StepCompleteWhen((_runOneStep OR _runAllSteps) AND _finishStep);

    IF _runOneStep THEN
        _runOneStep := FALSE;
        RETURN;
    END_IF
END_IF

IF SUPER^.Step(948, TRUE, 'Step number 948') THEN
    SUPER^.StepCompleteWhen((_runOneStep OR _runAllSteps) AND _finishStep);

    IF _runOneStep THEN
        _runOneStep := FALSE;
        RETURN;
    END_IF
END_IF

IF SUPER^.Step(949, TRUE, 'Step number 949') THEN
    SUPER^.StepCompleteWhen((_runOneStep OR _runAllSteps) AND _finishStep);

    IF _runOneStep THEN
        _runOneStep := FALSE;
        RETURN;
    END_IF
END_IF

IF SUPER^.Step(950, TRUE, 'Step number 950') THEN
    SUPER^.StepCompleteWhen((_runOneStep OR _runAllSteps) AND _finishStep);

    IF _runOneStep THEN
        _runOneStep := FALSE;
        RETURN;
    END_IF
END_IF

IF SUPER^.Step(951, TRUE, 'Step number 951') THEN
    SUPER^.StepCompleteWhen((_runOneStep OR _runAllSteps) AND _finishStep);

    IF _runOneStep THEN
        _runOneStep := FALSE;
        RETURN;
    END_IF
END_IF

IF SUPER^.Step(952, TRUE, 'Step number 952') THEN
    SUPER^.StepCompleteWhen((_runOneStep OR _runAllSteps) AND _finishStep);

    IF _runOneStep THEN
        _runOneStep := FALSE;
        RETURN;
    END_IF
END_IF

IF SUPER^.Step(953, TRUE, 'Step number 953') THEN
    SUPER^.StepCompleteWhen((_runOneStep OR _runAllSteps) AND _finishStep);

    IF _runOneStep THEN
        _runOneStep := FALSE;
        RETURN;
    END_IF
END_IF

IF SUPER^.Step(954, TRUE, 'Step number 954') THEN
    SUPER^.StepCompleteWhen((_runOneStep OR _runAllSteps) AND _finishStep);

    IF _runOneStep THEN
        _runOneStep := FALSE;
        RETURN;
    END_IF
END_IF

IF SUPER^.Step(955, TRUE, 'Step number 955') THEN
    SUPER^.StepCompleteWhen((_runOneStep OR _runAllSteps) AND _finishStep);

    IF _runOneStep THEN
        _runOneStep := FALSE;
        RETURN;
    END_IF
END_IF

IF SUPER^.Step(956, TRUE, 'Step number 956') THEN
    SUPER^.StepCompleteWhen((_runOneStep OR _runAllSteps) AND _finishStep);

    IF _runOneStep THEN
        _runOneStep := FALSE;
        RETURN;
    END_IF
END_IF

IF SUPER^.Step(957, TRUE, 'Step number 957') THEN
    SUPER^.StepCompleteWhen((_runOneStep OR _runAllSteps) AND _finishStep);

    IF _runOneStep THEN
        _runOneStep := FALSE;
        RETURN;
    END_IF
END_IF

IF SUPER^.Step(958, TRUE, 'Step number 958') THEN
    SUPER^.StepCompleteWhen((_runOneStep OR _runAllSteps) AND _finishStep);

    IF _runOneStep THEN
        _runOneStep := FALSE;
        RETURN;
    END_IF
END_IF

IF SUPER^.Step(959, TRUE, 'Step number 959') THEN
    SUPER^.StepCompleteWhen((_runOneStep OR _runAllSteps) AND _finishStep);

    IF _runOneStep THEN
        _runOneStep := FALSE;
        RETURN;
    END_IF
END_IF

IF SUPER^.Step(960, TRUE, 'Step number 960') THEN
    SUPER^.StepCompleteWhen((_runOneStep OR _runAllSteps) AND _finishStep);

    IF _runOneStep THEN
        _runOneStep := FALSE;
        RETURN;
    END_IF
END_IF

IF SUPER^.Step(961, TRUE, 'Step number 961') THEN
    SUPER^.StepCompleteWhen((_runOneStep OR _runAllSteps) AND _finishStep);

    IF _runOneStep THEN
        _runOneStep := FALSE;
        RETURN;
    END_IF
END_IF

IF SUPER^.Step(962, TRUE, 'Step number 962') THEN
    SUPER^.StepCompleteWhen((_runOneStep OR _runAllSteps) AND _finishStep);

    IF _runOneStep THEN
        _runOneStep := FALSE;
        RETURN;
    END_IF
END_IF

IF SUPER^.Step(963, TRUE, 'Step number 963') THEN
    SUPER^.StepCompleteWhen((_runOneStep OR _runAllSteps) AND _finishStep);

    IF _runOneStep THEN
        _runOneStep := FALSE;
        RETURN;
    END_IF
END_IF

IF SUPER^.Step(964, TRUE, 'Step number 964') THEN
    SUPER^.StepCompleteWhen((_runOneStep OR _runAllSteps) AND _finishStep);

    IF _runOneStep THEN
        _runOneStep := FALSE;
        RETURN;
    END_IF
END_IF

IF SUPER^.Step(965, TRUE, 'Step number 965') THEN
    SUPER^.StepCompleteWhen((_runOneStep OR _runAllSteps) AND _finishStep);

    IF _runOneStep THEN
        _runOneStep := FALSE;
        RETURN;
    END_IF
END_IF

IF SUPER^.Step(966, TRUE, 'Step number 966') THEN
    SUPER^.StepCompleteWhen((_runOneStep OR _runAllSteps) AND _finishStep);

    IF _runOneStep THEN
        _runOneStep := FALSE;
        RETURN;
    END_IF
END_IF

IF SUPER^.Step(967, TRUE, 'Step number 967') THEN
    SUPER^.StepCompleteWhen((_runOneStep OR _runAllSteps) AND _finishStep);

    IF _runOneStep THEN
        _runOneStep := FALSE;
        RETURN;
    END_IF
END_IF

IF SUPER^.Step(968, TRUE, 'Step number 968') THEN
    SUPER^.StepCompleteWhen((_runOneStep OR _runAllSteps) AND _finishStep);

    IF _runOneStep THEN
        _runOneStep := FALSE;
        RETURN;
    END_IF
END_IF

IF SUPER^.Step(969, TRUE, 'Step number 969') THEN
    SUPER^.StepCompleteWhen((_runOneStep OR _runAllSteps) AND _finishStep);

    IF _runOneStep THEN
        _runOneStep := FALSE;
        RETURN;
    END_IF
END_IF

IF SUPER^.Step(970, TRUE, 'Step number 970') THEN
    SUPER^.StepCompleteWhen((_runOneStep OR _runAllSteps) AND _finishStep);

    IF _runOneStep THEN
        _runOneStep := FALSE;
        RETURN;
    END_IF
END_IF

IF SUPER^.Step(971, TRUE, 'Step number 971') THEN
    SUPER^.StepCompleteWhen((_runOneStep OR _runAllSteps) AND _finishStep);

    IF _runOneStep THEN
        _runOneStep := FALSE;
        RETURN;
    END_IF
END_IF

IF SUPER^.Step(972, TRUE, 'Step number 972') THEN
    SUPER^.StepCompleteWhen((_runOneStep OR _runAllSteps) AND _finishStep);

    IF _runOneStep THEN
        _runOneStep := FALSE;
        RETURN;
    END_IF
END_IF

IF SUPER^.Step(973, TRUE, 'Step number 973') THEN
    SUPER^.StepCompleteWhen((_runOneStep OR _runAllSteps) AND _finishStep);

    IF _runOneStep THEN
        _runOneStep := FALSE;
        RETURN;
    END_IF
END_IF

IF SUPER^.Step(974, TRUE, 'Step number 974') THEN
    SUPER^.StepCompleteWhen((_runOneStep OR _runAllSteps) AND _finishStep);

    IF _runOneStep THEN
        _runOneStep := FALSE;
        RETURN;
    END_IF
END_IF

IF SUPER^.Step(975, TRUE, 'Step number 975') THEN
    SUPER^.StepCompleteWhen((_runOneStep OR _runAllSteps) AND _finishStep);

    IF _runOneStep THEN
        _runOneStep := FALSE;
        RETURN;
    END_IF
END_IF

IF SUPER^.Step(976, TRUE, 'Step number 976') THEN
    SUPER^.StepCompleteWhen((_runOneStep OR _runAllSteps) AND _finishStep);

    IF _runOneStep THEN
        _runOneStep := FALSE;
        RETURN;
    END_IF
END_IF

IF SUPER^.Step(977, TRUE, 'Step number 977') THEN
    SUPER^.StepCompleteWhen((_runOneStep OR _runAllSteps) AND _finishStep);

    IF _runOneStep THEN
        _runOneStep := FALSE;
        RETURN;
    END_IF
END_IF

IF SUPER^.Step(978, TRUE, 'Step number 978') THEN
    SUPER^.StepCompleteWhen((_runOneStep OR _runAllSteps) AND _finishStep);

    IF _runOneStep THEN
        _runOneStep := FALSE;
        RETURN;
    END_IF
END_IF

IF SUPER^.Step(979, TRUE, 'Step number 979') THEN
    SUPER^.StepCompleteWhen((_runOneStep OR _runAllSteps) AND _finishStep);

    IF _runOneStep THEN
        _runOneStep := FALSE;
        RETURN;
    END_IF
END_IF

IF SUPER^.Step(980, TRUE, 'Step number 980') THEN
    SUPER^.StepCompleteWhen((_runOneStep OR _runAllSteps) AND _finishStep);

    IF _runOneStep THEN
        _runOneStep := FALSE;
        RETURN;
    END_IF
END_IF

IF SUPER^.Step(981, TRUE, 'Step number 981') THEN
    SUPER^.StepCompleteWhen((_runOneStep OR _runAllSteps) AND _finishStep);

    IF _runOneStep THEN
        _runOneStep := FALSE;
        RETURN;
    END_IF
END_IF

IF SUPER^.Step(982, TRUE, 'Step number 982') THEN
    SUPER^.StepCompleteWhen((_runOneStep OR _runAllSteps) AND _finishStep);

    IF _runOneStep THEN
        _runOneStep := FALSE;
        RETURN;
    END_IF
END_IF

IF SUPER^.Step(983, TRUE, 'Step number 983') THEN
    SUPER^.StepCompleteWhen((_runOneStep OR _runAllSteps) AND _finishStep);

    IF _runOneStep THEN
        _runOneStep := FALSE;
        RETURN;
    END_IF
END_IF

IF SUPER^.Step(984, TRUE, 'Step number 984') THEN
    SUPER^.StepCompleteWhen((_runOneStep OR _runAllSteps) AND _finishStep);

    IF _runOneStep THEN
        _runOneStep := FALSE;
        RETURN;
    END_IF
END_IF

IF SUPER^.Step(985, TRUE, 'Step number 985') THEN
    SUPER^.StepCompleteWhen((_runOneStep OR _runAllSteps) AND _finishStep);

    IF _runOneStep THEN
        _runOneStep := FALSE;
        RETURN;
    END_IF
END_IF

IF SUPER^.Step(986, TRUE, 'Step number 986') THEN
    SUPER^.StepCompleteWhen((_runOneStep OR _runAllSteps) AND _finishStep);

    IF _runOneStep THEN
        _runOneStep := FALSE;
        RETURN;
    END_IF
END_IF

IF SUPER^.Step(987, TRUE, 'Step number 987') THEN
    SUPER^.StepCompleteWhen((_runOneStep OR _runAllSteps) AND _finishStep);

    IF _runOneStep THEN
        _runOneStep := FALSE;
        RETURN;
    END_IF
END_IF

IF SUPER^.Step(988, TRUE, 'Step number 988') THEN
    SUPER^.StepCompleteWhen((_runOneStep OR _runAllSteps) AND _finishStep);

    IF _runOneStep THEN
        _runOneStep := FALSE;
        RETURN;
    END_IF
END_IF

IF SUPER^.Step(989, TRUE, 'Step number 989') THEN
    SUPER^.StepCompleteWhen((_runOneStep OR _runAllSteps) AND _finishStep);

    IF _runOneStep THEN
        _runOneStep := FALSE;
        RETURN;
    END_IF
END_IF

IF SUPER^.Step(990, TRUE, 'Step number 990') THEN
    SUPER^.StepCompleteWhen((_runOneStep OR _runAllSteps) AND _finishStep);

    IF _runOneStep THEN
        _runOneStep := FALSE;
        RETURN;
    END_IF
END_IF

IF SUPER^.Step(991, TRUE, 'Step number 991') THEN
    SUPER^.StepCompleteWhen((_runOneStep OR _runAllSteps) AND _finishStep);

    IF _runOneStep THEN
        _runOneStep := FALSE;
        RETURN;
    END_IF
END_IF

IF SUPER^.Step(992, TRUE, 'Step number 992') THEN
    SUPER^.StepCompleteWhen((_runOneStep OR _runAllSteps) AND _finishStep);

    IF _runOneStep THEN
        _runOneStep := FALSE;
        RETURN;
    END_IF
END_IF

IF SUPER^.Step(993, TRUE, 'Step number 993') THEN
    SUPER^.StepCompleteWhen((_runOneStep OR _runAllSteps) AND _finishStep);

    IF _runOneStep THEN
        _runOneStep := FALSE;
        RETURN;
    END_IF
END_IF

IF SUPER^.Step(994, TRUE, 'Step number 994') THEN
    SUPER^.StepCompleteWhen((_runOneStep OR _runAllSteps) AND _finishStep);

    IF _runOneStep THEN
        _runOneStep := FALSE;
        RETURN;
    END_IF
END_IF

IF SUPER^.Step(995, TRUE, 'Step number 995') THEN
    SUPER^.StepCompleteWhen((_runOneStep OR _runAllSteps) AND _finishStep);

    IF _runOneStep THEN
        _runOneStep := FALSE;
        RETURN;
    END_IF
END_IF

IF SUPER^.Step(996, TRUE, 'Step number 996') THEN
    SUPER^.StepCompleteWhen((_runOneStep OR _runAllSteps) AND _finishStep);

    IF _runOneStep THEN
        _runOneStep := FALSE;
        RETURN;
    END_IF
END_IF

IF SUPER^.Step(997, TRUE, 'Step number 997') THEN
    SUPER^.StepCompleteWhen((_runOneStep OR _runAllSteps) AND _finishStep);

    IF _runOneStep THEN
        _runOneStep := FALSE;
        RETURN;
    END_IF
END_IF

IF SUPER^.Step(998, TRUE, 'Step number 998') THEN
    SUPER^.StepCompleteWhen((_runOneStep OR _runAllSteps) AND _finishStep);

    IF _runOneStep THEN
        _runOneStep := FALSE;
        RETURN;
    END_IF
END_IF

IF SUPER^.Step(999, TRUE, 'Step number 999') THEN
    SUPER^.StepCompleteWhen((_runOneStep OR _runAllSteps) AND _finishStep);

    IF _runOneStep THEN
        _runOneStep := FALSE;
        RETURN;
    END_IF
END_IF

IF SUPER^.Step(1000, TRUE, 'Step number 1000') THEN
    SUPER^.StepCompleteWhen((_runOneStep OR _runAllSteps) AND _finishStep);

    IF _runOneStep THEN
        _runOneStep := FALSE;
        RETURN;
    END_IF
END_IF

IF SUPER^.Step(1001, TRUE, 'Step number 1001') THEN
    SUPER^.StepCompleteWhen((_runOneStep OR _runAllSteps) AND _finishStep);

    IF _runOneStep THEN
        _runOneStep := FALSE;
        RETURN;
    END_IF
END_IF

IF SUPER^.Step(1002, TRUE, 'Step number 1002') THEN
    SUPER^.StepCompleteWhen((_runOneStep OR _runAllSteps) AND _finishStep);

    IF _runOneStep THEN
        _runOneStep := FALSE;
        RETURN;
    END_IF
END_IF

IF SUPER^.Step(1003, TRUE, 'Step number 1003') THEN
    SUPER^.StepCompleteWhen((_runOneStep OR _runAllSteps) AND _finishStep);

    IF _runOneStep THEN
        _runOneStep := FALSE;
        RETURN;
    END_IF
END_IF

IF SUPER^.Step(1004, TRUE, 'Step number 1004') THEN
    SUPER^.StepCompleteWhen((_runOneStep OR _runAllSteps) AND _finishStep);

    IF _runOneStep THEN
        _runOneStep := FALSE;
        RETURN;
    END_IF
END_IF

IF SUPER^.Step(1005, TRUE, 'Step number 1005') THEN
    SUPER^.StepCompleteWhen((_runOneStep OR _runAllSteps) AND _finishStep);

    IF _runOneStep THEN
        _runOneStep := FALSE;
        RETURN;
    END_IF
END_IF

IF SUPER^.Step(1006, TRUE, 'Step number 1006') THEN
    SUPER^.StepCompleteWhen((_runOneStep OR _runAllSteps) AND _finishStep);

    IF _runOneStep THEN
        _runOneStep := FALSE;
        RETURN;
    END_IF
END_IF

IF SUPER^.Step(1007, TRUE, 'Step number 1007') THEN
    SUPER^.StepCompleteWhen((_runOneStep OR _runAllSteps) AND _finishStep);

    IF _runOneStep THEN
        _runOneStep := FALSE;
        RETURN;
    END_IF
END_IF

IF SUPER^.Step(1008, TRUE, 'Step number 1008') THEN
    SUPER^.StepCompleteWhen((_runOneStep OR _runAllSteps) AND _finishStep);

    IF _runOneStep THEN
        _runOneStep := FALSE;
        RETURN;
    END_IF
END_IF

IF SUPER^.Step(1009, TRUE, 'Step number 1009') THEN
    SUPER^.StepCompleteWhen((_runOneStep OR _runAllSteps) AND _finishStep);

    IF _runOneStep THEN
        _runOneStep := FALSE;
        RETURN;
    END_IF
END_IF

IF SUPER^.Step(1010, TRUE, 'Step number 1010') THEN
    SUPER^.StepCompleteWhen((_runOneStep OR _runAllSteps) AND _finishStep);

    IF _runOneStep THEN
        _runOneStep := FALSE;
        RETURN;
    END_IF
END_IF

IF SUPER^.Step(1011, TRUE, 'Step number 1011') THEN
    SUPER^.StepCompleteWhen((_runOneStep OR _runAllSteps) AND _finishStep);

    IF _runOneStep THEN
        _runOneStep := FALSE;
        RETURN;
    END_IF
END_IF

IF SUPER^.Step(1012, TRUE, 'Step number 1012') THEN
    SUPER^.StepCompleteWhen((_runOneStep OR _runAllSteps) AND _finishStep);

    IF _runOneStep THEN
        _runOneStep := FALSE;
        RETURN;
    END_IF
END_IF

IF SUPER^.Step(1013, TRUE, 'Step number 1013') THEN
    SUPER^.StepCompleteWhen((_runOneStep OR _runAllSteps) AND _finishStep);

    IF _runOneStep THEN
        _runOneStep := FALSE;
        RETURN;
    END_IF
END_IF

IF SUPER^.Step(1014, TRUE, 'Step number 1014') THEN
    SUPER^.StepCompleteWhen((_runOneStep OR _runAllSteps) AND _finishStep);

    IF _runOneStep THEN
        _runOneStep := FALSE;
        RETURN;
    END_IF
END_IF

IF SUPER^.Step(1015, TRUE, 'Step number 1015') THEN
    SUPER^.StepCompleteWhen((_runOneStep OR _runAllSteps) AND _finishStep);

    IF _runOneStep THEN
        _runOneStep := FALSE;
        RETURN;
    END_IF
END_IF

IF SUPER^.Step(1016, TRUE, 'Step number 1016') THEN
    SUPER^.StepCompleteWhen((_runOneStep OR _runAllSteps) AND _finishStep);

    IF _runOneStep THEN
        _runOneStep := FALSE;
        RETURN;
    END_IF
END_IF

IF SUPER^.Step(1017, TRUE, 'Step number 1017') THEN
    SUPER^.StepCompleteWhen((_runOneStep OR _runAllSteps) AND _finishStep);

    IF _runOneStep THEN
        _runOneStep := FALSE;
        RETURN;
    END_IF
END_IF

IF SUPER^.Step(1018, TRUE, 'Step number 1018') THEN
    SUPER^.StepCompleteWhen((_runOneStep OR _runAllSteps) AND _finishStep);

    IF _runOneStep THEN
        _runOneStep := FALSE;
        RETURN;
    END_IF
END_IF

IF SUPER^.Step(1019, TRUE, 'Step number 1019') THEN
    SUPER^.StepCompleteWhen((_runOneStep OR _runAllSteps) AND _finishStep);

    IF _runOneStep THEN
        _runOneStep := FALSE;
        RETURN;
    END_IF
END_IF

IF SUPER^.Step(1020, TRUE, 'Step number 1020') THEN
    SUPER^.StepCompleteWhen((_runOneStep OR _runAllSteps) AND _finishStep);

    IF _runOneStep THEN
        _runOneStep := FALSE;
        RETURN;
    END_IF
END_IF

IF SUPER^.Step(1021, TRUE, 'Step number 1021') THEN
    SUPER^.StepCompleteWhen((_runOneStep OR _runAllSteps) AND _finishStep);

    IF _runOneStep THEN
        _runOneStep := FALSE;
        RETURN;
    END_IF
END_IF

IF SUPER^.Step(1022, TRUE, 'Step number 1022') THEN
    SUPER^.StepCompleteWhen((_runOneStep OR _runAllSteps) AND _finishStep);

    IF _runOneStep THEN
        _runOneStep := FALSE;
        RETURN;
    END_IF
END_IF

IF SUPER^.Step(1023, TRUE, 'Step number 1023') THEN
    SUPER^.StepCompleteWhen((_runOneStep OR _runAllSteps) AND _finishStep);

    IF _runOneStep THEN
        _runOneStep := FALSE;
        RETURN;
    END_IF
END_IF

//******************************************************************
IF SUPER^.Step(_stepId, _enabled, _stepDescription) THEN
    SUPER^.StepCompleteWhen((_runOneStep OR _runAllSteps) AND _finishStep);

    IF _runOneStep THEN
        _runOneStep := FALSE;
        RETURN;
    END_IF
END_IF
END_METHOD

METHOD MAIN_CommentOutPartOfRunningSequencer 
VAR 
	i : INT;
END_VAR
IF _sequenceRun =1 THEN
	IF Step(0, TRUE, 'Step 0') THEN
	   StepCompleteWhen(TRUE);
	END_IF

	IF Step(1, TRUE, 'Step 1') THEN
	   StepCompleteWhen(TRUE);
	END_IF

	IF Step(2, TRUE, 'Step 2') THEN
	   StepCompleteWhen(TRUE);
	END_IF

	IF Step(3, TRUE, 'Step 3') THEN
			StepCompleteWhen(FALSE);
	END_IF
	
	FOR i := 4 TO _totalStepNumber-2 DO
		IF Step(i, TRUE, CONCAT('Step ', INT_TO_STRING(i))) THEN
			StepCompleteWhen(FALSE);
		END_IF
	END_FOR
	
	IF Step(_totalStepNumber - 1, TRUE, CONCAT('Step ', INT_TO_STRING(_totalStepNumber - 1))) THEN
	  _SequenceComplete();
	END_IF
END_IF

IF _sequenceRun >=2 THEN
	IF Step(0, TRUE, 'Step 0') THEN
	   StepCompleteWhen(TRUE);
	END_IF

//	IF Step(1, TRUE, 'Step 1') THEN
//	   StepCompleteWhen(TRUE);
//	END_IF

//	IF Step(2, TRUE, 'Step 2') THEN
//	   StepCompleteWhen(TRUE);
//	END_IF

	IF Step(3, TRUE, 'Step 3') THEN
	   StepCompleteWhen(FALSE);
	END_IF
	
	FOR i := 4 TO _totalStepNumber-2 DO
		IF Step(i, TRUE, CONCAT('Step ', INT_TO_STRING(i))) THEN
			StepCompleteWhen(FALSE);
		END_IF
	END_FOR
	
	IF Step(_totalStepNumber - 1, TRUE, CONCAT('Step ', INT_TO_STRING(_totalStepNumber - 1))) THEN
	  _SequenceComplete();
	END_IF
END_IF
END_METHOD

METHOD MAIN_ExecutionInOnePLCcycle 
VAR 
	i : INT;
END_VAR
FOR i := 0 TO _totalStepNumber-2 DO
    IF Step(i, TRUE, CONCAT('Step ', INT_TO_STRING(i))) THEN
        StepCompleteWhen(TRUE);
    END_IF
END_FOR

IF Step(_totalStepNumber - 1, TRUE, CONCAT('Step ', INT_TO_STRING(_totalStepNumber - 1))) THEN
   	_SequenceComplete();
END_IF
END_METHOD

METHOD MAIN_MaxStepId 
VAR 
	i : INT;
END_VAR
FOR i := 0 TO _totalStepNumber-1 DO
    IF Step(i, TRUE, CONCAT('Step ', INT_TO_STRING(i))) THEN
        StepCompleteWhen(_finishStep);
    END_IF
END_FOR
IF Step(_stepId, TRUE, CONCAT('Step ', INT_TO_STRING(_stepId))) THEN
    StepCompleteWhen(TRUE);
END_IF
END_METHOD

METHOD MAIN_MinStepId 
VAR 
	i : INT;
END_VAR
IF Step(_stepId, TRUE, CONCAT('Step ', INT_TO_STRING(_stepId))) THEN
    StepCompleteWhen(TRUE);
END_IF

FOR i := 1 TO _totalStepNumber-1 DO
    IF Step(i, TRUE, CONCAT('Step ', INT_TO_STRING(i))) THEN
        StepCompleteWhen(_finishStep);
    END_IF
END_FOR
END_METHOD

METHOD MAIN_NumberOfStepsCount 
VAR 
	i : INT;
END_VAR
IF Step(0, TRUE, 'Step 0') THEN
    StepCompleteWhen(TRUE);
END_IF

FOR i := 1 TO _totalStepNumber - 1 DO
    IF Step(i, TRUE, CONCAT('Step ', INT_TO_STRING(i))) THEN
        StepCompleteWhen(_finishStep);
    END_IF
END_FOR
END_METHOD

METHOD MAIN_OnStateChangeWhenChangingModes 
VAR 
	i : INT;
END_VAR
IF _sequenceRun <= _cyclicCycles OR _sequenceRun > _cyclicCycles + _stepInEvents + 1 THEN
    SetCyclicMode();

    FOR i := 0 TO _totalStepNumber - 2 DO
        IF Step(i, TRUE, CONCAT('Step ', INT_TO_STRING(i))) THEN
            _StepCompleteWhen(TRUE);
        END_IF
    END_FOR

    IF Step(_totalStepNumber - 1, TRUE, CONCAT('Step ', INT_TO_STRING(_totalStepNumber - 1))) THEN
        CompleteSequence();
		_sequenceCycles := _sequenceCycles + 1;
    END_IF
END_IF
IF _sequenceRun = _cyclicCycles+1 THEN
    SetStepMode();
	Step(0,FALSE,'');	
END_IF
IF _sequenceRun > _cyclicCycles+1  AND _sequenceRun <= _cyclicCycles + _stepInEvents +1 THEN
    SetStepMode();
	_StepIn();
    FOR i := 0 TO _totalStepNumber - 2 DO
        IF Step(i, TRUE, CONCAT('Step ', INT_TO_STRING(i))) THEN
            _StepCompleteWhen(TRUE);
        END_IF
    END_FOR

    IF Step(_totalStepNumber - 1, TRUE, CONCAT('Step ', INT_TO_STRING(_totalStepNumber - 1))) THEN
        CompleteSequence();
		_sequenceCycles := _sequenceCycles + 1;
    END_IF
END_IF
END_METHOD

METHOD MAIN_RequestStep 
VAR 
	i : INT;
END_VAR
IF _sequenceRun =1 THEN
	FOR i := -5 TO -1 DO
		IF Step(i, TRUE, CONCAT('Step ', INT_TO_STRING(i))) THEN
			StepCompleteWhen(TRUE);
		END_IF
	END_FOR
	
	IF Step(0, TRUE, 'Step 0') THEN
		RequestStep(-5);
	END_IF
	
	FOR i := 1 TO 5 DO
		IF Step(i, TRUE, CONCAT('Step ', INT_TO_STRING(i))) THEN
			StepCompleteWhen(TRUE);
		END_IF
	END_FOR
END_IF

IF _sequenceRun =2 THEN
	FOR i := -5 TO 5 DO
		IF Step(i, TRUE, CONCAT('Step ', INT_TO_STRING(i))) THEN
			StepCompleteWhen(FALSE);
		END_IF
	END_FOR
END_IF

IF _sequenceRun =3 THEN
	IF Step(-5, TRUE, 'Step -5') THEN
		RequestStep(0);
	END_IF

	FOR i := -4 TO 5 DO
		IF Step(i, TRUE, CONCAT('Step ', INT_TO_STRING(i))) THEN
			StepCompleteWhen(FALSE);
		END_IF
	END_FOR
END_IF
END_METHOD

METHOD MAIN_RequestStepFromHigherToLower 
VAR 
	i : INT;
END_VAR
IF _sequenceRun = 1 THEN
    FOR i := 0 TO _reqStep + 4 DO
        IF Step(i, TRUE, CONCAT('Step ', INT_TO_STRING(i))) THEN
            StepCompleteWhen(TRUE);
        END_IF
    END_FOR

    FOR i := _reqStep + 5 TO _totalStepNumber - 2 DO
        Step(i, TRUE, CONCAT('Step ', INT_TO_STRING(i)));
    END_FOR

    RequestStep(_reqStep);

    IF Step(_totalStepNumber - 1, TRUE, CONCAT('Step ', INT_TO_STRING(_totalStepNumber - 1))) THEN
        _SequenceComplete();
    END_IF
END_IF

IF _sequenceRun = 2 THEN
    FOR i := 0 TO _totalStepNumber - 2 DO
        Step(i, TRUE, CONCAT('Step ', INT_TO_STRING(i)));
    END_FOR

    IF Step(_totalStepNumber - 1, TRUE, CONCAT('Step ', INT_TO_STRING(_totalStepNumber - 1))) THEN
        _SequenceComplete();
    END_IF
END_IF
END_METHOD

METHOD MAIN_RequestStepFromLowerToHigher 
VAR 
	i : INT;
END_VAR
IF _sequenceRun = 1 THEN
    IF Step(0, TRUE, 'Step 0') THEN
        StepCompleteWhen(TRUE);
    END_IF

    FOR i := 1 TO _totalStepNumber - 2 DO
        Step(i, TRUE, CONCAT('Step ', INT_TO_STRING(i)));
    END_FOR

    IF Step(_totalStepNumber - 1, TRUE, CONCAT('Step ', INT_TO_STRING(_totalStepNumber - 1))) THEN
        _SequenceComplete();
    END_IF
END_IF

IF _sequenceRun = 2 THEN
    IF Step(0, TRUE, 'Step 0') THEN
        StepCompleteWhen(TRUE);
    END_IF

    RequestStep(_reqStep);

    FOR i := 1 TO _totalStepNumber - 2 DO
        Step(i, TRUE, CONCAT('Step ', INT_TO_STRING(i)));
    END_FOR

    IF Step(_totalStepNumber - 1, TRUE, CONCAT('Step ', INT_TO_STRING(_totalStepNumber - 1))) THEN
        _SequenceComplete();
    END_IF
END_IF
END_METHOD

METHOD MAIN_RequestStepToFirstStepWithStepId0 
VAR 
	i : INT;
END_VAR
FOR i := 0 TO 4 DO
    IF Step(i, TRUE, CONCAT('Step ', INT_TO_STRING(i))) THEN
        StepCompleteWhen(_finishStep);
    END_IF
END_FOR

IF Step(5, TRUE, 'Step 5') THEN
    RequestStep(0);
END_IF

FOR i := 6 TO _totalStepNumber DO
    IF Step(i, TRUE, CONCAT('Step ', INT_TO_STRING(i))) THEN
        StepCompleteWhen(_finishStep);
    END_IF
END_FOR
END_METHOD

METHOD MAIN_RequestStepToNotExistingStep 
VAR 
	i : INT;
END_VAR
IF _sequenceRun = 1 THEN
    RequestStep(_reqStepNotExists);

    FOR i := 0 TO _totalStepNumber - 2 DO
        Step(i, TRUE, CONCAT('Step ', INT_TO_STRING(i)));
    END_FOR

    IF Step(_totalStepNumber - 1, TRUE, CONCAT('Step ', INT_TO_STRING(_totalStepNumber - 1))) THEN
        _SequenceComplete();
    END_IF
END_IF

IF _sequenceRun >= 2 THEN
    FOR i := 0 TO _totalStepNumber - 2 DO
        Step(i, TRUE, CONCAT('Step ', INT_TO_STRING(i)));
    END_FOR

    IF Step(_totalStepNumber - 1, TRUE, CONCAT('Step ', INT_TO_STRING(_totalStepNumber - 1))) THEN
        _SequenceComplete();
    END_IF
END_IF
END_METHOD

METHOD MAIN_RequestStepWhilePreviousRequestStepHasNotBeenYetProcessed 
VAR 
	i : INT;
END_VAR
FOR i := 0 TO _reqStep + 4 DO
    IF Step(i, TRUE, CONCAT('Step ', INT_TO_STRING(i))) THEN
        StepCompleteWhen(TRUE);
    END_IF
END_FOR

RequestStep(_reqStep);

FOR i := _reqStep + 5 TO _totalStepNumber - 2 DO
    Step(i, TRUE, CONCAT('Step ', INT_TO_STRING(i)));
END_FOR

RequestStep(_reqStep + 10);

IF Step(_totalStepNumber - 1, TRUE, CONCAT('Step ', INT_TO_STRING(_totalStepNumber - 1))) THEN
    _SequenceComplete();
END_IF
END_METHOD

METHOD MAIN_RestoreChildBetweenSteps 
VAR 
	i : INT;
	_childState : INT;
END_VAR
FOR i := 0 TO _totalStepNumber-2 DO
    IF Step(i, TRUE, CONCAT('Step ', INT_TO_STRING(i))) THEN
		_childState := _myTcoChildState.State;
		_myTcoChildState.ChangeState(_myTcoChildState._requestedState);
        StepCompleteWhen(TRUE);
    END_IF
END_FOR

IF Step(_totalStepNumber - 1, TRUE, CONCAT('Step ', INT_TO_STRING(_totalStepNumber - 1))) THEN
   	_SequenceComplete();
END_IF
END_METHOD

METHOD MAIN_SetStepMode 
VAR 
	i : INT;
END_VAR
IF _sequenceRun = 1 THEN
    IF Step(0, TRUE, 'Initial step') THEN
        StepCompleteWhen(TRUE);
    END_IF

    FOR i := 1 TO _totalStepNumber - 2 DO
        Step(i, TRUE, CONCAT('Step ', INT_TO_STRING(i)));
    END_FOR

    IF Step(_totalStepNumber - 1, TRUE, CONCAT('Step ', INT_TO_STRING(_totalStepNumber - 1))) THEN
        _SequenceComplete();
    END_IF
END_IF

IF _sequenceRun =4 THEN
    IF Step(0, TRUE, 'Initial step') THEN
        StepCompleteWhen(TRUE);
    END_IF

    FOR i := 1 TO _totalStepNumber - 2 DO
        IF Step(i, TRUE, CONCAT('Step ', INT_TO_STRING(i))) THEN
	        StepCompleteWhen(TRUE);
		END_IF
    END_FOR

    IF Step(_totalStepNumber - 1, TRUE, CONCAT('Step ', INT_TO_STRING(_totalStepNumber - 1))) THEN
        _SequenceComplete();
    END_IF
END_IF
END_METHOD

METHOD MAIN_StepMode 
VAR 
	i : INT;
END_VAR
IF _sequenceRun = 1 THEN
    IF Step(0, TRUE, 'Initial step') THEN
        StepCompleteWhen(TRUE);
    END_IF

    FOR i := 1 TO _totalStepNumber - 2 DO
        Step(i, TRUE, CONCAT('Step ', INT_TO_STRING(i)));
    END_FOR

    IF Step(_totalStepNumber - 1, TRUE, CONCAT('Step ', INT_TO_STRING(_totalStepNumber - 1))) THEN
        _SequenceComplete();
    END_IF
END_IF

IF _sequenceRun > 1 THEN
    _StepIn();

    IF Step(0, TRUE, 'Initial step') THEN
        StepCompleteWhen(TRUE);
    END_IF

    FOR i := 1 TO _totalStepNumber - 2 DO
        IF Step(i, TRUE, CONCAT('Step ', INT_TO_STRING(i))) THEN
            StepCompleteWhen(TRUE);
        END_IF
    END_FOR

    IF Step(_totalStepNumber - 1, TRUE, CONCAT('Step ', INT_TO_STRING(_totalStepNumber - 1))) THEN
        _SequenceComplete();
    END_IF
END_IF
END_METHOD

METHOD MAIN_StepModeChangeStepIdDuringExecution 
VAR 
	i : INT;
END_VAR
IF _sequenceRun = 1 THEN
    IF _currentStep.Status = 20 THEN
       _StepIn();
    END_IF

    // Step 0
    IF Step(0, TRUE, 'Step 0') THEN
        StepCompleteWhen(TRUE);
    END_IF

    // Step 1
    IF Step(1, TRUE, 'Step 1') THEN
        StepCompleteWhen(TRUE);
    END_IF

    // Step 2
    IF Step(2, TRUE, 'Step 2') THEN
        StepCompleteWhen(TRUE);
    END_IF

    // Step 3
    IF Step(3, TRUE, 'Step 3') THEN
        StepCompleteWhen(FALSE);
    END_IF

    FOR i := 4 TO _totalStepNumber - 2 DO
        Step(i, TRUE, CONCAT('Step  ', INT_TO_STRING(i)));
    END_FOR

    IF Step(_totalStepNumber - 1, TRUE, CONCAT('Step  ', INT_TO_STRING(_totalStepNumber - 1))) THEN
        _SequenceComplete();
    END_IF
END_IF
IF _sequenceRun = 2 THEN
    IF _currentStep.Status = 20 THEN
       _StepIn();
    END_IF

    // Step 0
    IF Step(0, TRUE, 'Step 0') THEN
        StepCompleteWhen(TRUE);
    END_IF

    // Step 1
    IF Step(1, TRUE, 'Step 1') THEN
        StepCompleteWhen(TRUE);
    END_IF

    // Step 2
    IF Step(2, TRUE, 'Step 2') THEN
        StepCompleteWhen(TRUE);
    END_IF

    // Step 3
    IF Step(5, TRUE, 'Step 3') THEN
        StepCompleteWhen(FALSE);
    END_IF

    FOR i := 4 TO _totalStepNumber - 2 DO
        Step(i, TRUE, CONCAT('Step  ', INT_TO_STRING(i)));
    END_FOR

    IF Step(_totalStepNumber - 1, TRUE, CONCAT('Step  ', INT_TO_STRING(_totalStepNumber - 1))) THEN
        _SequenceComplete();
    END_IF
END_IF
END_METHOD

METHOD MAIN_StepModeChangeStepOrder 
VAR 
	i : INT;
END_VAR
IF _sequenceRun <= _totalStepNumber + 1 THEN
    IF _currentStep.Status = 20 THEN
       _StepIn();
    END_IF

    // Step 0
    IF Step(0, TRUE, 'Step 0') THEN
        StepCompleteWhen(TRUE);
    END_IF

    // Step 1
    IF Step(1, TRUE, 'Step 1') THEN
        StepCompleteWhen(TRUE);
    END_IF

    // Step 2
    IF Step(2, TRUE, 'Step 2') THEN
        StepCompleteWhen(TRUE);
    END_IF

    // Step 3
    IF Step(3, TRUE, 'Step 3') THEN
        StepCompleteWhen(FALSE);
    END_IF

    FOR i := 4 TO _totalStepNumber - 2 DO
        Step(i, TRUE, CONCAT('Step  ', INT_TO_STRING(i)));
    END_FOR

    IF Step(_totalStepNumber-1, TRUE, CONCAT('Step  ', INT_TO_STRING(_totalStepNumber-1))) THEN
        _SequenceComplete();
    END_IF
END_IF
IF _sequenceRun = _totalStepNumber + 2 THEN
    IF _currentStep.Status = 20 THEN
       _StepIn();
    END_IF

    // Step 0
    IF Step(0, TRUE, 'Step 0') THEN
        StepCompleteWhen(TRUE);
    END_IF

    // Step 1
    IF Step(1, TRUE, 'Step 1') THEN
        StepCompleteWhen(TRUE);
    END_IF

    // Step 3
    IF Step(3, TRUE, 'Step 3') THEN
        StepCompleteWhen(FALSE);
    END_IF

    // Step 2
    IF Step(2, TRUE, 'Step 2') THEN
        StepCompleteWhen(TRUE);
    END_IF

    FOR i := 4 TO _totalStepNumber - 2 DO
        Step(i, TRUE, CONCAT('Step  ', INT_TO_STRING(i)));
    END_FOR

    IF Step(_totalStepNumber-1, TRUE, CONCAT('Step  ', INT_TO_STRING(_totalStepNumber-1))) THEN
        _SequenceComplete();
    END_IF
END_IF
END_METHOD

METHOD MAIN_StepModeCommentOutPartOfRunningSequencer 
VAR 
	i : INT;
END_VAR
IF _sequenceRun =1 THEN
    IF (_currentStep.Status = 20) THEN
        _StepIn();
    END_IF

	IF Step(0, TRUE, 'Step 0') THEN
	   StepCompleteWhen(TRUE);
	END_IF

	IF Step(1, TRUE, 'Step 1') THEN
	   StepCompleteWhen(TRUE);
	END_IF

	IF Step(2, TRUE, 'Step 2') THEN
	   StepCompleteWhen(TRUE);
	END_IF

	IF Step(3, TRUE, 'Step 3') THEN
			StepCompleteWhen(FALSE);
	END_IF
	
	FOR i := 4 TO _totalStepNumber-2 DO
		IF Step(i, TRUE, CONCAT('Step ', INT_TO_STRING(i))) THEN
			StepCompleteWhen(FALSE);
		END_IF
	END_FOR
	
	IF Step(_totalStepNumber-1, TRUE, CONCAT('Step ', INT_TO_STRING(_totalStepNumber-1))) THEN
	  _SequenceComplete();
	END_IF
END_IF

IF _sequenceRun >=2 THEN
    IF (_currentStep.Status = 20) THEN
        _StepIn();
    END_IF

	IF Step(0, TRUE, 'Step 0') THEN
	   StepCompleteWhen(TRUE);
	END_IF

//	IF Step(1, TRUE, 'Step 1') THEN
//	   StepCompleteWhen(TRUE);
//	END_IF

//	IF Step(2, TRUE, 'Step 2') THEN
//	   StepCompleteWhen(TRUE);
//	END_IF

	IF Step(3, TRUE, 'Step 3') THEN
	   StepCompleteWhen(FALSE);
	END_IF
	
	FOR i := 4 TO _totalStepNumber-2 DO
		IF Step(i, TRUE, CONCAT('Step ', INT_TO_STRING(i))) THEN
			StepCompleteWhen(FALSE);
		END_IF
	END_FOR
	
	IF Step(_totalStepNumber-1, TRUE, CONCAT('Step ', INT_TO_STRING(_totalStepNumber-1))) THEN
	  _SequenceComplete();
	END_IF
END_IF
END_METHOD

METHOD MAIN_StepModeDisabledStep 
VAR 
	i : INT;
END_VAR
IF _sequenceRun = 1 THEN
    FOR i := 0 TO _totalStepNumber-1 DO
        Step(i, TRUE, CONCAT('Step ', INT_TO_STRING(i)));
    END_FOR
END_IF

IF _sequenceRun = 2 OR _sequenceRun = 3 THEN
    IF _sequenceRun = 2 THEN
        _StepIn();
    END_IF

    IF Step(0, TRUE, 'Step 0') THEN
        StepCompleteWhen(TRUE);
    END_IF

    FOR i := 1 TO _totalStepNumber - 2 DO
        Step(i, TRUE, CONCAT('Step ', INT_TO_STRING(i)));
    END_FOR

    IF Step(_totalStepNumber-1, TRUE, CONCAT('Step ', INT_TO_STRING(_totalStepNumber-1))) THEN
        CompleteSequence();
    END_IF
END_IF

IF _sequenceRun = 4 THEN
    IF Step(0, TRUE, 'Step 0') THEN
        StepCompleteWhen(TRUE);
    END_IF

    IF Step(1, FALSE, 'Step 1') THEN
        StepCompleteWhen(TRUE);
    END_IF

    FOR i := 2 TO _totalStepNumber - 2 DO
        Step(i, TRUE, CONCAT('Step ', INT_TO_STRING(i)));
    END_FOR

    IF Step(_totalStepNumber-1, TRUE, CONCAT('Step ', INT_TO_STRING(_totalStepNumber-1))) THEN
        CompleteSequence();
    END_IF
END_IF

IF _sequenceRun >= 5 THEN
    _StepIn();

    IF Step(0, TRUE, 'Step 0') THEN
        StepCompleteWhen(TRUE);
    END_IF

    IF Step(1, FALSE, 'Step 1') THEN
        StepCompleteWhen(TRUE);
    END_IF

    FOR i := 2 TO _totalStepNumber - 2 DO
        Step(i, TRUE, CONCAT('Step ', INT_TO_STRING(i)));
    END_FOR

    IF Step(_totalStepNumber-1, TRUE, CONCAT('Step ', INT_TO_STRING(_totalStepNumber-1))) THEN
        CompleteSequence();
    END_IF
END_IF
END_METHOD

METHOD MAIN_StepModeRequestStepFromHigherToLower 
VAR 
	i : INT;
END_VAR
IF _sequenceRun <=_reqStep + 5 THEN
    FOR i := 0 TO _reqStep + 4 DO
       _StepIn();
        IF Step(i, TRUE, CONCAT('Step ', INT_TO_STRING(i))) THEN
            StepCompleteWhen(TRUE);
        END_IF
    END_FOR

    FOR i := _reqStep + 5 TO _totalStepNumber - 2 DO
       _StepIn();
        Step(i, TRUE, CONCAT('Step ', INT_TO_STRING(i)));
    END_FOR

    IF Step(_totalStepNumber-1, TRUE, CONCAT('Step ', INT_TO_STRING(_totalStepNumber-1))) THEN
        _SequenceComplete();
    END_IF
END_IF

IF _sequenceRun =_reqStep + 6 THEN
    FOR i := 0 TO _reqStep + 4 DO
       _StepIn();
        IF Step(i, TRUE, CONCAT('Step ', INT_TO_STRING(i))) THEN
            StepCompleteWhen(TRUE);
        END_IF
    END_FOR

    FOR i := _reqStep + 5 TO _totalStepNumber - 2 DO
       _StepIn();
        Step(i, TRUE, CONCAT('Step ', INT_TO_STRING(i)));
    END_FOR

    RequestStep(_reqStep);

    IF Step(_totalStepNumber-1, TRUE, CONCAT('Step ', INT_TO_STRING(_totalStepNumber-1))) THEN
        _SequenceComplete();
    END_IF
END_IF

IF _sequenceRun >=_reqStep + 7 THEN
    FOR i := 0 TO _totalStepNumber - 2 DO
       _StepIn();
        Step(i, TRUE, CONCAT('Step ', INT_TO_STRING(i)));
    END_FOR

    IF Step(_totalStepNumber-1, TRUE, CONCAT('Step ', INT_TO_STRING(_totalStepNumber-1))) THEN
        _SequenceComplete();
    END_IF
END_IF
END_METHOD

METHOD MAIN_StepModeRequestStepFromLowerToHigher 
VAR 
	i : INT;
END_VAR
IF _sequenceRun = 1 THEN
    IF _currentStep.Status = 20 THEN
       _StepIn();
    END_IF
    IF Step(0, TRUE, 'Step 0') THEN
        StepCompleteWhen(TRUE);
    END_IF

    FOR i := 1 TO _totalStepNumber - 2 DO
        Step(i, TRUE, CONCAT('Step ', INT_TO_STRING(i)));
    END_FOR

    IF Step(_totalStepNumber-1, TRUE, CONCAT('Step ', INT_TO_STRING(_totalStepNumber-1))) THEN
        _SequenceComplete();
    END_IF
END_IF

IF _sequenceRun = 2 THEN
    IF _currentStep.Status = 20 THEN
       _StepIn();
    END_IF
    IF Step(0, TRUE, 'Step 0') THEN
        StepCompleteWhen(TRUE);
    END_IF

    RequestStep(_reqStep);

    FOR i := 1 TO _totalStepNumber - 2 DO
        Step(i, TRUE, CONCAT('Step ', INT_TO_STRING(i)));
    END_FOR

    IF Step(_totalStepNumber-1, TRUE, CONCAT('Step ', INT_TO_STRING(_totalStepNumber-1))) THEN
        _SequenceComplete();
    END_IF
END_IF
END_METHOD

METHOD MAIN_StepModeStepBackwardFromRunningStep 
VAR 
	i : INT;
END_VAR
IF _sequenceRun = 1 THEN
    _StepIn();
END_IF

IF _sequenceRun = 11 THEN
    _StepBackward();
END_IF

Step(0, TRUE, 'Step 0');
Step(1, TRUE, 'Step 1');

IF Step(2, TRUE, 'Step 2') THEN
    _StepCompleteWhen(_sequenceRun >= 20);
END_IF

IF Step(3, TRUE, 'Step 3') THEN
    _StepCompleteWhen(_sequenceRun >= 20);
END_IF

FOR i := 4 TO _totalStepNumber - 2 DO
    Step(i, TRUE, CONCAT('Step ', INT_TO_STRING(i)));
END_FOR

IF Step(_totalStepNumber-1, TRUE, CONCAT('Step ', INT_TO_STRING(_totalStepNumber-1))) THEN
    CompleteSequence();
END_IF
END_METHOD

METHOD MAIN_StepModeStepForwardBackward 
VAR 
	i : INT;
END_VAR
IF _sequenceRun = 1 THEN
    FOR i := 0 TO _totalStepNumber - 2 DO
        Step(i, TRUE, CONCAT('Step ', INT_TO_STRING(i)));
    END_FOR

    IF Step(_totalStepNumber - 1, TRUE, CONCAT('Step ', INT_TO_STRING(_totalStepNumber - 1))) THEN
        CompleteSequence();
    END_IF
END_IF

IF _sequenceRun = 2 THEN
    _StepIn();

    IF Step(0, TRUE, 'Step 0') THEN
        StepCompleteWhen(TRUE);
    END_IF

    FOR i := 1 TO _totalStepNumber - 2 DO
        Step(i, TRUE, CONCAT('Step ', INT_TO_STRING(i)));
    END_FOR

    IF Step(_totalStepNumber - 1, TRUE, CONCAT('Step ', INT_TO_STRING(_totalStepNumber- 1))) THEN
        CompleteSequence();
    END_IF
END_IF

IF _sequenceRun = 3 OR _sequenceRun = 5 THEN
    _StepForward();

    IF Step(0, TRUE, 'Step 0') THEN
        StepCompleteWhen(TRUE);
    END_IF

    FOR i := 1 TO _totalStepNumber - 2 DO
        Step(i, TRUE, CONCAT('Step ', INT_TO_STRING(i)));
    END_FOR

    IF Step(_totalStepNumber - 1, TRUE, CONCAT('Step ', INT_TO_STRING(_totalStepNumber - 1))) THEN
        CompleteSequence();
    END_IF
END_IF

IF _sequenceRun = 4 THEN
    RequestStep(_totalStepNumber -1);

    IF Step(0, TRUE, 'Step 0') THEN
        StepCompleteWhen(TRUE);
    END_IF

    FOR i := 1 TO _totalStepNumber - 2 DO
        Step(i, TRUE, CONCAT('Step ', INT_TO_STRING(i)));
    END_FOR

    IF Step(_totalStepNumber - 1, TRUE, CONCAT('Step ', INT_TO_STRING(_totalStepNumber - 1))) THEN
        CompleteSequence();
    END_IF
END_IF

IF _sequenceRun = 6 OR _sequenceRun = 8 OR _sequenceRun = 9 THEN
    _StepBackward();

    IF Step(0, TRUE, 'Step 0') THEN
        StepCompleteWhen(TRUE);
    END_IF

    FOR i := 1 TO _totalStepNumber - 2 DO
        Step(i, TRUE, CONCAT('Step ', INT_TO_STRING(i)));
    END_FOR

    IF Step(_totalStepNumber-1, TRUE, CONCAT('Step ', INT_TO_STRING(_totalStepNumber-1))) THEN
        CompleteSequence();
    END_IF
END_IF

IF _sequenceRun = 7 THEN
    RequestStep(1);

    IF Step(0, TRUE, 'Step 0') THEN
        StepCompleteWhen(TRUE);
    END_IF

    FOR i := 1 TO _totalStepNumber - 2 DO
        Step(i, TRUE, CONCAT('Step ', INT_TO_STRING(i)));
    END_FOR

    IF Step(_totalStepNumber-1, TRUE, CONCAT('Step ', INT_TO_STRING(_totalStepNumber-1))) THEN
        CompleteSequence();
    END_IF
END_IF
END_METHOD

METHOD MAIN_StepModeStepForwardFromRunningStep 
VAR 
	i : INT;
END_VAR
IF _sequenceRun = 1 THEN
    _StepIn();
END_IF

IF _sequenceRun = 11 THEN
    _StepForward();
END_IF

Step(0, TRUE, 'Step 0');
Step(1, TRUE, 'Step 1');

IF Step(2, TRUE, 'Step 2') THEN
    _StepCompleteWhen(_sequenceRun >= 20);
END_IF

IF Step(3, TRUE, 'Step 3') THEN
    _StepCompleteWhen(_sequenceRun >= 20);
END_IF

FOR i := 4 TO _totalStepNumber - 2 DO
    Step(i, TRUE, CONCAT('Step ', INT_TO_STRING(i)));
END_FOR

IF Step(_totalStepNumber-1, TRUE, CONCAT('Step ', INT_TO_STRING(_totalStepNumber-1))) THEN
    CompleteSequence();
END_IF
END_METHOD

METHOD MAIN_StepModeStepIn 
VAR 
	i : INT;
END_VAR
IF _sequenceRun = 1 THEN
    IF Step(0, TRUE, 'Initial step') THEN
        StepCompleteWhen(TRUE);
    END_IF

    FOR i := 1 TO _totalStepNumber - 2 DO
        Step(i, TRUE, CONCAT('Step ', INT_TO_STRING(i)));
    END_FOR

    IF Step(_totalStepNumber-1, TRUE, CONCAT('Step ', INT_TO_STRING(_totalStepNumber-1))) THEN
        _SequenceComplete();
    END_IF
END_IF

IF _sequenceRun > 1 THEN
    IF _currentStep.Status = 20 THEN
       _StepIn();
    END_IF

    // Step 0
    IF Step(0, TRUE, 'Step 0') THEN
        StepCompleteWhen(TRUE);
    END_IF

    // Step 1
    IF Step(1, TRUE, 'Step 1') THEN
        StepCompleteWhen(TRUE);
    END_IF

    // Step 2
    IF Step(2, TRUE, 'Step 2') THEN
        StepCompleteWhen(TRUE);
    END_IF

    // Step 3
    IF Step(3, TRUE, 'Step 3') THEN
        StepCompleteWhen(FALSE);
    END_IF

    FOR i := 4 TO _totalStepNumber - 2 DO
        Step(i, TRUE, CONCAT('Step  ', INT_TO_STRING(i)));
    END_FOR

    IF Step(_totalStepNumber-1, TRUE, CONCAT('Step  ', INT_TO_STRING(_totalStepNumber-1))) THEN
        _SequenceComplete();
    END_IF
END_IF
END_METHOD

METHOD MAIN_StepModeStepInDetailed 
VAR 
	i : INT;
END_VAR
IF _sequenceRun = 1 OR _sequenceRun = 5 THEN
    FOR i := 0 TO _totalStepNumber - 2 DO
        Step(i, TRUE, CONCAT('Step ', INT_TO_STRING(i)));
    END_FOR

    IF Step(_totalStepNumber - 1, TRUE, CONCAT('Step ', INT_TO_STRING(_totalStepNumber - 1))) THEN
        CompleteSequence();
    END_IF
END_IF

IF _sequenceRun = 2 THEN
    _StepIn();

    IF Step(0, TRUE, 'Step 0') THEN
        StepCompleteWhen(TRUE);
    END_IF

    FOR i := 1 TO _totalStepNumber - 2 DO
        Step(i, TRUE, CONCAT('Step ', INT_TO_STRING(i)));
    END_FOR

    IF Step(_totalStepNumber - 1, TRUE, CONCAT('Step ', INT_TO_STRING(_totalStepNumber - 1))) THEN
        CompleteSequence();
    END_IF
END_IF

IF _sequenceRun = 3 OR _sequenceRun = 4 THEN
    _StepIn();

    IF Step(0, TRUE, 'Step 0') THEN
        StepCompleteWhen(TRUE);
    END_IF

    IF Step(1, TRUE, 'Step 1') THEN
        RequestStep(_totalStepNumber - 1);
    END_IF

    FOR i := 2 TO _totalStepNumber - 2 DO
        Step(i, TRUE, CONCAT('Step ', INT_TO_STRING(i)));
    END_FOR

    IF Step(_totalStepNumber - 1, TRUE, CONCAT('Step ', INT_TO_STRING(_totalStepNumber - 1))) THEN
        CompleteSequence();
    END_IF
END_IF
END_METHOD

METHOD MAIN_StepModeUncommentPartOfRunningSequencer 
VAR 
	i : INT;
END_VAR
IF _sequenceRun = 1 THEN
    IF (_currentStep.Status = 20) THEN
        _StepIn();
    END_IF

    IF Step(0, TRUE, 'Step 0') THEN
        StepCompleteWhen(TRUE);
    END_IF

    //	IF Step(1, TRUE, 'Step 1') THEN
    //	   StepCompleteWhen(TRUE);
    //	END_IF
    //	IF Step(2, TRUE, 'Step 2') THEN
    //	   StepCompleteWhen(TRUE);
    //	END_IF
    IF Step(3, TRUE, 'Step 3') THEN
        StepCompleteWhen(FALSE);
    END_IF

    FOR i := 4 TO _totalStepNumber - 2 DO
        IF Step(i, TRUE, CONCAT('Step ', INT_TO_STRING(i))) THEN
            StepCompleteWhen(FALSE);
        END_IF
    END_FOR

    IF Step(_totalStepNumber-1, TRUE, CONCAT('Step ', INT_TO_STRING(_totalStepNumber-1))) THEN
        _SequenceComplete();
    END_IF
END_IF

IF _sequenceRun = 2 THEN
    IF (_currentStep.Status = 20) THEN
        _StepIn();
    END_IF

    IF Step(0, TRUE, 'Step 0') THEN
        StepCompleteWhen(TRUE);
    END_IF

    IF Step(1, TRUE, 'Step 1') THEN
        StepCompleteWhen(TRUE);
    END_IF

    IF Step(2, TRUE, 'Step 2') THEN
        StepCompleteWhen(TRUE);
    END_IF

    IF Step(3, TRUE, 'Step 3') THEN
        StepCompleteWhen(FALSE);
    END_IF

    FOR i := 4 TO _totalStepNumber - 2 DO
        IF Step(i, TRUE, CONCAT('Step ', INT_TO_STRING(i))) THEN
            StepCompleteWhen(FALSE);
        END_IF
    END_FOR

    IF Step(_totalStepNumber-1, TRUE, CONCAT('Step ', INT_TO_STRING(_totalStepNumber-1))) THEN
        _SequenceComplete();
    END_IF
END_IF
END_METHOD

METHOD MAIN_SwitchStepModeOnDuringStepExecution 
VAR 
	i : INT;
END_VAR
IF _sequenceRun = 1 THEN
    IF Step(0, TRUE, 'Step 0') THEN
        StepCompleteWhen(TRUE);
    END_IF

    IF Step(1, TRUE, 'Step 1') THEN
        StepCompleteWhen(FALSE);
    END_IF

    FOR i := 2 TO _totalStepNumber - 2 DO
        Step(i, TRUE, CONCAT('Step ', INT_TO_STRING(i)));
    END_FOR

    IF Step(_totalStepNumber-1, TRUE, CONCAT('Step ', INT_TO_STRING(_totalStepNumber-1))) THEN
        CompleteSequence();
    END_IF
END_IF

IF _sequenceRun > 1 THEN
    IF Step(0, TRUE, 'Step 0') THEN
        StepCompleteWhen(TRUE);
    END_IF

    IF Step(1, TRUE, 'Step 1') THEN
		IF _sequenceRun >=5 THEN
			SetStepMode();
		END_IF
        StepCompleteWhen(_sequenceRun >=10);
    END_IF

    FOR i := 2 TO _totalStepNumber - 2 DO
        Step(i, TRUE, CONCAT('Step ', INT_TO_STRING(i)));
    END_FOR

    IF Step(_totalStepNumber-1, TRUE, CONCAT('Step ', INT_TO_STRING(_totalStepNumber-1))) THEN
        CompleteSequence();
    END_IF
END_IF
END_METHOD

METHOD MAIN_SwitchStepModeStepOffFromReadyToRun 
VAR 
	i : INT;
END_VAR
SetCyclicMode();
Step(0, TRUE, 'Step 0');
Step(1, TRUE, 'Step 1');

IF Step(2, TRUE, 'Step 2') THEN
    _StepCompleteWhen(_sequenceRun >= 20);
END_IF

IF Step(3, TRUE, 'Step 3') THEN
    _StepCompleteWhen(_sequenceRun >= 20);
END_IF

FOR i := 4 TO _totalStepNumber - 2 DO
    Step(i, TRUE, CONCAT('Step ', INT_TO_STRING(i)));
END_FOR

IF Step(_totalStepNumber-1, TRUE, CONCAT('Step ', INT_TO_STRING(_totalStepNumber-1))) THEN
    CompleteSequence();
END_IF
END_METHOD

METHOD MAIN_SwitchStepModeStepOffFromRunning 
VAR 
	i : INT;
END_VAR
SetCyclicMode();
Step(0, TRUE, 'Step 0');
Step(1, TRUE, 'Step 1');

IF Step(2, TRUE, 'Step 2') THEN
    _StepCompleteWhen(_sequenceRun >= 20);
END_IF

IF Step(3, TRUE, 'Step 3') THEN
    _StepCompleteWhen(_sequenceRun >= 20);
END_IF

FOR i := 4 TO _totalStepNumber - 2 DO
    Step(i, TRUE, CONCAT('Step ', INT_TO_STRING(i)));
END_FOR

IF Step(_totalStepNumber-1, TRUE, CONCAT('Step ', INT_TO_STRING(_totalStepNumber-1))) THEN
    CompleteSequence();
END_IF
END_METHOD

METHOD MAIN_SwitchStepModeStepOnFromRunning 
VAR 
	i : INT;
END_VAR
SetStepMode();
Step(0, TRUE, 'Step 0');
Step(1, TRUE, 'Step 1');

IF Step(2, TRUE, 'Step 2') THEN
    _StepCompleteWhen(_sequenceRun >= 20);
END_IF

IF Step(3, TRUE, 'Step 3') THEN
    _StepCompleteWhen(_sequenceRun >= 20);
END_IF

FOR i := 4 TO _totalStepNumber - 2 DO
    Step(i, TRUE, CONCAT('Step ', INT_TO_STRING(i)));
END_FOR

IF Step(_totalStepNumber-1, TRUE, CONCAT('Step ', INT_TO_STRING(_totalStepNumber-1))) THEN
    CompleteSequence();
END_IF
END_METHOD

METHOD MAIN_UncommentPartOfRunningSequencer 
VAR 
	i : INT;
END_VAR
IF _sequenceRun =1 THEN
	IF Step(0, TRUE, 'Step 0') THEN
	   StepCompleteWhen(TRUE);
	END_IF

//	IF Step(1, TRUE, 'Step 1') THEN
//	   StepCompleteWhen(TRUE);
//	END_IF

//	IF Step(2, TRUE, 'Step 2') THEN
//	   StepCompleteWhen(TRUE);
//	END_IF

	IF Step(3, TRUE, 'Step 3') THEN
	   StepCompleteWhen(FALSE);
	END_IF
	
	FOR i := 4 TO _totalStepNumber-2 DO
		IF Step(i, TRUE, CONCAT('Step ', INT_TO_STRING(i))) THEN
			StepCompleteWhen(FALSE);
		END_IF
	END_FOR
	
	IF Step(_totalStepNumber-1, TRUE, CONCAT('Step ', INT_TO_STRING(_totalStepNumber-1))) THEN
	  _SequenceComplete();
	END_IF
END_IF

IF _sequenceRun =2 THEN
	IF Step(0, TRUE, 'Step 0') THEN
	   StepCompleteWhen(TRUE);
	END_IF

	IF Step(1, TRUE, 'Step 1') THEN
	   StepCompleteWhen(TRUE);
	END_IF

	IF Step(2, TRUE, 'Step 2') THEN
	   StepCompleteWhen(TRUE);
	END_IF

	IF Step(3, TRUE, 'Step 3') THEN
			StepCompleteWhen(FALSE);
	END_IF
	
	FOR i := 4 TO _totalStepNumber-2 DO
		IF Step(i, TRUE, CONCAT('Step ', INT_TO_STRING(i))) THEN
			StepCompleteWhen(FALSE);
		END_IF
	END_FOR
	
	IF Step(_totalStepNumber-1, TRUE, CONCAT('Step ', INT_TO_STRING(_totalStepNumber-1))) THEN
	  _SequenceComplete();
	END_IF
END_IF
END_METHOD

METHOD PROTECTED OnRestore
_restoreCycleCount := _restoreCycleCount + 1;
END_METHOD

METHOD PROTECTED OnSequenceCompleted
_onSequenceCompleteCount := _onSequenceCompleteCount + 1;
END_METHOD

METHOD PROTECTED OnSequencerError
VAR_INPUT
	inErrorId : eSequencerError;
END_VAR
CASE inErrorId OF
	eSequencerError.noError :
		_onSequencerErrorCount := _onSequencerErrorCount + 0;
	eSequencerError.NotUniqueStepId :
		_onSequencerErrorCount := _onSequencerErrorCount + 10;
	eSequencerError.StepIdHasBeenChanged :
		_onSequencerErrorCount := _onSequencerErrorCount + 20;
	eSequencerError.OrderOfTheStepHasBeenChanged :
		_onSequencerErrorCount := _onSequencerErrorCount + 40;
	eSequencerError.StepWithRequestedIdDoesNotExists :
		_onSequencerErrorCount := _onSequencerErrorCount + 50;
	eSequencerError.MultipleRequestStepMethodCall :
		_onSequencerErrorCount := _onSequencerErrorCount + 60;
	eSequencerError.StepIdTooLow :
		_onSequencerErrorCount := _onSequencerErrorCount + 70;
	eSequencerError.StepIdTooHigh :
		_onSequencerErrorCount := _onSequencerErrorCount + 80;
	ELSE
		_onSequencerErrorCount := _onSequencerErrorCount + 0;
END_CASE
END_METHOD

METHOD PROTECTED OnStateChange
VAR_INPUT
	PreviousState	: INT;
	NewState 		: INT;
END_VAR
THIS^._onStateChangeCount := THIS^._onStateChangeCount + 1;

_stateChangeFrom := PreviousState;
_stateChangeTo := NewState;

IF _callRestoreInOnStateChange THEN
	Restore();
END_IF
END_METHOD

METHOD PROTECTED OnStepCompleted
_onCompleteStepCount := _onCompleteStepCount + 1;
END_METHOD

PROPERTY PostOpenRequestStepCycle : UINT
GET
PostOpenRequestStepCycle := _postOpenRequestStepCycle;
END_GET
SET
_postOpenRequestStepCycle := PostOpenRequestStepCycle;
END_SET
END_PROPERTY

PROPERTY PreCloseRequestStepCycle : UINT
GET
PreCloseRequestStepCycle := _preCloseRequestStepCycle;
END_GET
SET
_preCloseRequestStepCycle := PreCloseRequestStepCycle;
END_SET
END_PROPERTY

PROPERTY ReqStep : INT
GET
ReqStep := _reqStep;
END_GET
SET
_reqStep := ReqStep;
END_SET
END_PROPERTY

PROPERTY ReqStepNotExists : INT
GET
ReqStepNotExists := _reqStepNotExists;
END_GET
SET
_reqStepNotExists:=ReqStepNotExists;
END_SET
END_PROPERTY

PROPERTY INTERNAL RequestStepCycle : UINT
GET
RequestStepCycle := _requestStepCycle;
END_GET
SET
_requestStepCycle := RequestStepCycle;
END_SET
END_PROPERTY

PROPERTY RunAllSteps : BOOL
GET
RunAllSteps := _runAllSteps;
END_GET
SET
_runAllSteps := RunAllSteps;
END_SET
END_PROPERTY

PROPERTY RunOneStep : BOOL
GET
RunOneStep := _runOneStep;
END_GET
SET
_runOneStep := RunOneStep;
END_SET
END_PROPERTY

{attribute 'TcRpcEnable'}
METHOD SaveNumberOfStepsInSequence
_numberOfSteps := THIS^._numberOfStepsInSequence;
_previousNumberOfSteps	:= THIS^._previousNumberOfStepsInSequence;
END_METHOD

PROPERTY SequenceCycles : UINT
GET
SequenceCycles := _sequenceCycles;
END_GET
SET
_sequenceCycles := SequenceCycles;
END_SET
END_PROPERTY

METHOD INTERNAL SequencerClose
SUPER^._Close();
END_METHOD

METHOD INTERNAL SequencerOpen
SUPER^._Open();
END_METHOD

PROPERTY SequenceRun : ULINT
GET
SequenceRun := _sequenceRun;
END_GET
SET
_sequenceRun:=SequenceRun;
END_SET
END_PROPERTY

{attribute 'TcRpcEnable'}
METHOD INTERNAL SetChildState 
VAR_INPUT
	inState			:	INT;
END_VAR
THIS^._myTcoChildState.ChangeState(inState);
END_METHOD

{attribute 'TcRpcEnable'}
METHOD INTERNAL SetCurrentStep 
VAR_INPUT
	inStepID 			:	INT;
	inStepDescription	:	STRING(254);
END_VAR
THIS^._currentStep.ID			:=	inStepID;
THIS^._currentStep.Description	:=	inStepDescription;
END_METHOD

{attribute 'TcRpcEnable'}
METHOD SetCurrentStepToErrorState : BOOL
_currentStep.Status := TcoCore.eStepStatus.Error;

SetCurrentStepToErrorState := _currentStep.Status = TcoCore.eStepStatus.Error;
END_METHOD

METHOD SetCyclicMode : BOOL
ModeController.Mode := eSequencerMode.CyclicMode;

SetCyclicMode := ModeController.Mode = eSequencerMode.CyclicMode;
END_METHOD

{attribute 'TcRpcEnable'}
METHOD SetInvalidMode : BOOL
ModeController.Mode := eSequencerMode.Invalid;

SetInvalidMode := ModeController.Mode = eSequencerMode.Invalid;
END_METHOD

METHOD INTERNAL SetNumberOfSteps 
VAR_INPUT
	inNumberOfSteps : UINT;
END_VAR
_stepCounter 						:=	inNumberOfSteps;
_numberOfStepsInSequence			:=	inNumberOfSteps;
_previousNumberOfStepsInSequence 	:=	inNumberOfSteps;
END_METHOD

METHOD INTERNAL SetSequenceAsChecked
_stepIDUniquenessChecked := TRUE;
_StepIdUniquenessControlState := eStepIdUniquenessControlState.Done;
END_METHOD

METHOD INTERNAL SetSequenceAsNotChecked
_stepIDUniquenessChecked := FALSE;
_StepIdUniquenessControlState := eStepIdUniquenessControlState.NotYetStarted;
END_METHOD

METHOD SetStepMode : BOOL
ModeController.Mode := eSequencerMode.StepMode;

SetStepMode := ModeController.Mode = eSequencerMode.StepMode;
END_METHOD

{attribute 'TcRpcEnable'}
METHOD INTERNAL SetupChildRequestedState 
VAR_INPUT
	inState			:	INT;
END_VAR
THIS^._myTcoChildState.RequestedState:=inState;
END_METHOD

PROPERTY StepDescription : STRING(254);
GET
StepDescription := _stepDescription;
END_GET
SET
_stepDescription := StepDescription;
END_SET
END_PROPERTY

PROPERTY StepId : INT
GET
StepId := _stepId;
END_GET
SET
_stepId := StepId;
END_SET
END_PROPERTY

PROPERTY StepInEvents : UINT
GET
StepInEvents := _stepInEvents;
END_GET
SET
_stepInEvents := StepInEvents;
END_SET
END_PROPERTY

PROPERTY TcoSequencerTest : eTcoSequencerTests
GET
TcoSequencerTest := _tcoSequencerTest;
END_GET
SET
_tcoSequencerTest := TcoSequencerTest;
END_SET
END_PROPERTY

PROPERTY TotalStepNumber : UINT
GET
TotalStepNumber := _totalStepNumber;
END_GET
SET
_totalStepNumber := TotalStepNumber;
END_SET
END_PROPERTY

END_FUNCTION_BLOCK

// ---- Tests/TcoSequencer/PlcExecuted/TcoSequencerTestChildState.TcPOU
FUNCTION_BLOCK TcoSequencerTestChildState EXTENDS TcoCore.TcoState
VAR
	_requestedState : UINT;
	_requestedStateCount :ULINT;
	_restoreCount :ULINT;
END_VAR

(*~
	<docu>
		<summary>
			This method is called on each change of the <c>State</c>. This method could be overloaded and custom code should be placed here.	
		</summary>			
	</docu>	
~*)
METHOD PROTECTED OnStateChange
VAR_INPUT
	PreviousState	: INT;
	NewState 		: INT;
END_VAR
IF NewState =  _requestedState THEN
	_requestedStateCount := _requestedStateCount + 1;
END_IF

IF NewState =  -1 THEN
	_restoreCount := _restoreCount + 1;
END_IF
END_METHOD

PROPERTY RequestedState : UINT
GET
RequestedState := _requestedState;
END_GET
SET
_requestedState := RequestedState;
END_SET
END_PROPERTY

END_FUNCTION_BLOCK

// ---- Tests/TcoSequence/PlcExecuted/TcoSequenceTestContext.TcPOU
FUNCTION_BLOCK TcoSequenceTestContext EXTENDS TcoCore._internals_TcoContext
VAR
    _sut_A : TcoSequenceTestType(THIS^, eRestoreMode.AutoRestoreMembers);
    _sut_N : TcoSequenceTestType(THIS^, eRestoreMode.None);

    _elapsedTimeETA : TIME;
    _elapsedTime : TIME;
    _runElapsedTimer : BOOL;
    _elapsedTimeTimer : Tc2_Standard.TON;

	_runOneStep							:	BOOL;
	_runAllSteps						:	BOOL;
	_finishStep							:	BOOL;
	_stepId								:	INT;
	_enabled							:	BOOL;
	_stepDescription					:	STRING(254);	
	_currentStepId						:	INT;
	_currentStepDescription				:	STRING(254);
    _totalStepNumber : UINT;
	_reqStep : INT;
    _reqStepNotExists : INT;

    _done : BOOL;
    _arranged : BOOL;
	_startCycles			:	ULINT;
	_endCycles				:	ULINT;	
	_myIdentity				:	ULINT;	
	_initReqStepCycle		:	UINT;
	_cycles					:	UINT;
	_cyclicCycles :	UINT;
    _stepInEvents :	UINT;

	//eTcoSequenceTests.FreshStateEntry:
	FreshStateEntry_counter : INT;
	FreshStateEntry_enter_and_leave_must_be_true : BOOL;
	FreshStateEntry_enter_and_two_cycles_on_first_must_be_true : BOOL;
	FreshStateEntry_enter_and_two_cycles_on_second_must_be_false : BOOL;
	FreshStateEntry_on_multiple_calls_but_not_first_must_be_false : BOOL;	
	FreshStateEntry_on_request_step_single_call_must_be_true : BOOL;	
END_VAR

{attribute 'TcRpcEnable'}
METHOD _ClearPlcCycleCounter
ClearPlcCycleCounter();
END_METHOD

METHOD PROTECTED Main
VAR
	i:INT;
END_VAR
_elapsedTimeTimer(IN := _runElapsedTimer, PT := _elapsedTimeETA);

CASE _testId OF
	eTcoSequenceTests.Initialize:
		_sut_A.Restore();
		_sut_N.Restore();
		FreshStateEntry_counter := 0;		
		FreshStateEntry_enter_and_leave_must_be_true := FALSE;
		FreshStateEntry_enter_and_two_cycles_on_first_must_be_true := FALSE;
		FreshStateEntry_enter_and_two_cycles_on_second_must_be_false := TRUE;
		FreshStateEntry_on_multiple_calls_but_not_first_must_be_false := TRUE;	
    {region "CallSequencerBodiesOnly"}
    eTcoSequenceTests.CallSequencerBodiesOnly:
        _sut_A.TcoSequencerTest := eTcoSequenceTests.CallSequencerBodiesOnly;
        _sut_N.TcoSequencerTest := eTcoSequenceTests.CallSequencerBodiesOnly;
        _sut_A._RunExecutionSubstitute();
        _sut_N._RunExecutionSubstitute();
    {endregion}
    {region "RestoreSequencers"}
    eTcoSequenceTests.RestoreSequencers:
        IF NOT _arranged THEN
            _sut_A.Restore();
            _sut_N.Restore();
            _arranged := _sut_A._restoringSequence AND _sut_N._restoringSequence;
        END_IF

        IF _arranged AND NOT _done THEN
            _sut_A.TcoSequencerTest := eTcoSequenceTests.RestoreSequencers;
            _sut_N.TcoSequencerTest := eTcoSequenceTests.RestoreSequencers;
            _sut_A._RunExecutionSubstitute();
            _sut_N._RunExecutionSubstitute();

            _done :=
                NOT _sut_A._restoringSequence AND NOT _sut_N._restoringSequence AND NOT _sut_A._sequencerHasError AND NOT _sut_N._sequencerHasError;
        END_IF

        ProbeDoneWhen(_done);
    {endregion}
    {region "T500_NumberOfStepsCount"}
    eTcoSequenceTests.NumberOfStepsCount:
        IF NOT _arranged THEN
            _sut_A.SetCyclicMode(); //Set sequencer into the cyclic mode
            _sut_N.SetCyclicMode(); //Set sequencer into the cyclic mode
            _sut_A.SetSequenceAsChecked(); //Set sequence as checked, so no StepID uniqueness is performed on next sequence execution
            _sut_N.SetSequenceAsChecked(); //Set sequence as checked, so no StepID uniqueness is performed on next sequence execution
            _sut_A.ClearNumberOfSteps(); //Clear internal flow step counters, so number of steps is going to be counted again on next sequence run
            _sut_N.ClearNumberOfSteps(); //Clear internal flow step counters, so number of steps is going to be counted again on next sequence run

            _sut_A.SetCurrentStep(_currentStepId,
                _currentStepDescription); //Set the StepId so as the StepDescription to the current step of the sequencer

            _sut_N.SetCurrentStep(_currentStepId,
                _currentStepDescription); //Set the StepId so as the StepDescription to the current step of the sequencer

            _sut_A.SaveNumberOfStepsInSequence();
            _sut_N.SaveNumberOfStepsInSequence();
            _sut_A.TcoSequencerTest := eTcoSequenceTests.NumberOfStepsCount;
            _sut_N.TcoSequencerTest := eTcoSequenceTests.NumberOfStepsCount;
            _sut_A.TotalStepNumber := _totalStepNumber;
            _sut_N.TotalStepNumber := _totalStepNumber;
            _sut_A.FinishStep := FALSE;
            _sut_N.FinishStep := FALSE;
            _arranged := TRUE;
            RETURN;
        END_IF

        IF NOT _done THEN
            _sut_A._RunExecutionSubstitute();
            _sut_N._RunExecutionSubstitute();
            _sut_A.SaveNumberOfStepsInSequence();
            _sut_N.SaveNumberOfStepsInSequence();
            _done := TRUE;
        END_IF

        IF _done THEN
            ProbeDoneWhen(_done);
        END_IF
    {endregion}
    {region "T501_ExecutionInOnePLCcycle"}
    eTcoSequenceTests.ExecutionInOnePLCcycle:
        _sut_A.TcoSequencerTest := eTcoSequenceTests.ExecutionInOnePLCcycle;
        _sut_N.TcoSequencerTest := eTcoSequenceTests.ExecutionInOnePLCcycle;
        _sut_A.SetCyclicMode(); //Set sequencer into the cyclic mode
        _sut_N.SetCyclicMode(); //Set sequencer into the cyclic mode
        _sut_A.TotalStepNumber := _totalStepNumber;
        _sut_N.TotalStepNumber := _totalStepNumber;
        _sut_A._RunExecutionSubstitute();
        _sut_N._RunExecutionSubstitute();
        _done := TRUE;
        ProbeDoneWhen(_done);
    {endregion}
    {region "T502_OnStepCompleted"}
    eTcoSequenceTests.OnStepCompleted:
        _sut_A.TcoSequencerTest := eTcoSequenceTests.OnStepCompleted;
        _sut_N.TcoSequencerTest := eTcoSequenceTests.OnStepCompleted;
        _sut_A.TotalStepNumber := _totalStepNumber;
        _sut_N.TotalStepNumber := _totalStepNumber;
        _sut_A._RunExecutionSubstitute();
        _sut_N._RunExecutionSubstitute();
        _sut_A.SaveNumberOfStepsInSequence();
        _sut_N.SaveNumberOfStepsInSequence();
        _done := TRUE;
        ProbeDoneWhen(_done);
    {endregion}
    {region "T503_OnSequenceCompleted"}
    eTcoSequenceTests.OnSequenceCompleted:
        _sut_A.TcoSequencerTest := eTcoSequenceTests.OnSequenceCompleted;
        _sut_N.TcoSequencerTest := eTcoSequenceTests.OnSequenceCompleted;
        _sut_A.TotalStepNumber := _totalStepNumber;
        _sut_N.TotalStepNumber := _totalStepNumber;
        _sut_A._RunExecutionSubstitute();
        _sut_N._RunExecutionSubstitute();
        _done := TRUE;
        ProbeDoneWhen(_done);
    {endregion}
    {region "T504_RestoreChildBetweenSteps"}
    eTcoSequenceTests.RestoreChildBetweenSteps:
        IF NOT _arranged THEN
            _sut_A.TcoSequencerTest := eTcoSequenceTests.RestoreChildBetweenSteps;
            _sut_N.TcoSequencerTest := eTcoSequenceTests.RestoreChildBetweenSteps;
            _sut_A.TotalStepNumber := _totalStepNumber;
            _sut_N.TotalStepNumber := _totalStepNumber;
            _arranged := TRUE;
            RETURN;
        END_IF;

